(* IEC 61131-3 sources: brOscatLib/oscatBasic (part 2) *)

(* ---- DWORD_TO_STRB.st ---- *)
FUNCTION DWORD_TO_STRB
    (*http://www.oscat.de/images/OSCATBasic/oscat_basic333_en.pdf#page=153*)
    (* pointer für die ausgabe ermitteln *)
    pt ACCESS ADR(RETVAL);
    (* die 8 ausgabecharacter ermitteln und schreiben *)
    FOR i := 1 TO 32 DO
    	pt:= USINT_TO_BYTE(BOOL_TO_USINT(IN.31) + 48);
    	IN := SHL(IN,1);
    	pt ACCESS (ADR(pt) + 1);
    END_FOR

    (* der ausgabestring muss nochg mit 0 abgeschlossen werden *)
    pt := 0;
    DWORD_TO_STRB := TRUE;

    (* revision history
    hm		9.6.2007	rev 1.0
    	original version

    hm		15.dec 2007	rev 1.1
    	changed code for better performance

    hm	29. mar. 2008	rev 1.2
    	changed STRING to STRING(32)

    hm	20. jun. 2008	rev 1.3
    	performance improvement

    *)

END_FUNCTION

(* ---- DWORD_TO_STRF.st ---- *)
FUNCTION DWORD_TO_STRF
    (*http://www.oscat.de/images/OSCATBasic/oscat_basic333_en.pdf#page=154*)
    (* limit N to max 20 characters *)
    (* convert dword to string first and cut to length N *)
    temp := DWORD_TO_STRING(IN);
    FIX(temp,LIMIT(0,N,20),48,1, RETVAL);
    DWORD_TO_STRF := TRUE;

    (* revision history
    hm	26. jan.2007	rev 1.0
    	original version

    hm	29. mar. 2008	rev 1.1
    	changed STRING to STRING(20)
    	limit the output string to max 20 digits
    *)

END_FUNCTION

(* ---- DWORD_TO_STRH.st ---- *)
FUNCTION DWORD_TO_STRH
    (*http://www.oscat.de/images/OSCATBasic/oscat_basic333_en.pdf#page=154*)
    (* read output adress to pointer *)
    pt ACCESS (ADR(DWORD_TO_STRH) + 8);
    (* wirte the closing byte for the string *)
    pt:= 0;

    (* write the 8 hex characters backwards *)
    FOR i := 1 TO 8 DO;
    	(* decrement the pointer *)
    	pt ACCESS (ADR(pt) - 1);
    	(* read the lowest order hex value *)
    	temp := DWORD_TO_BYTE(IN AND 16#0000000F);
        intTemp := BYTE_TO_USINT(temp);
    	(* convert value to hex character *)
    	IF intTemp <= 9 THEN temp := USINT_TO_BYTE(intTemp + 48); ELSE temp := USINT_TO_BYTE(intTemp + 55); END_IF
    	(* write character to output string *)
    	pt := temp;
    	(* shift IN for nect hex character *)
    	IN := SHR(IN,4);
    END_FOR

    (* code beofre rev 1.2
    FOR i := 1 TO 8 DO
    	X := DWORD_TO_BYTE(IN AND 2#1111);
    	IF X <= 9 THEN X := X + 48; ELSE X := X + 55; END_IF
    	Cx := CHR(X);
    	temp := CONCAT(Cx, temp);
    	IN := SHR(IN,4);
    END_FOR
    DWORD_TO_STRH := temp;
    *)

    (* revision history
    hm	9. jun. 2007	rev 1.0
    	original version

    hm	11. sep. 2007	rev 1.1
    	changed coding for compatibility with twincat, concat cannot support a function as an argument.

    hm	15. dec. 2007	rev 1.2
    	changed code for better performance

    hm	29. mar. 2008	rev 1.3
    	changed STRING to STRING(8)

    *)

END_FUNCTION

(* ---- EASTER.st ---- *)
FUNCTION EASTER
    (*http://www.oscat.de/images/OSCATBasic/oscat_basic333_en.pdf#page=122*)
    b := (204 - 11 * (YEAR MOD 19)) MOD 30;
    IF b > 27 THEN b := b - 1; END_IF
    c := (YEAR + SHR(YEAR,2) + b - 13) MOD 7;
    oday := 28 + b - c;
    IF oday > 33 THEN
    	EASTER := SET_DATE(YEAR, 4, oday - 31);
    ELSE
    	EASTER := SET_DATE(YEAR, 3, oday);
    END_IF

    (* alternativer algorithmus ueber das pasah fest
    execution time roughly 200us
    Der sog. Passah-Vollmond wird berechnet, in dem das Jahr durch 19 ge-
    teilt wird und der Rest mit der folgenden Tabelle verglichen wird:

        0: Apr 14       5: Apr 18      10: Mrz 25      15: Mrz 30
        1: Apr 03       6: Apr 08      11: Apr 13      16: Apr 17
        2: Mrz 23       7: Mrz 28      12: Apr 02      17: Apr 07
        3: Apr 11       8: Apr 16      13: Mrz 22      18: Mrz 27
        4: Mrz 31       9: Apr 05      14: Apr 10

    Faellt dieses Datum auf einen Sonntag, ist Ostern der naechste Sonntag!

    Beispiel: 1992 MOD 19 = 16, daraus folgt 17.04., der naechste Sonntag
              ist dann der 19. April (Ostersonntag)
    *)

    (* this algorithm is 180 us
    a := YEAR MOD 19;
    b := YEAR / 100;
    c := YEAR MOD 100;
    d := b / 4;
    e := b MOD 4;
    f := (b + 8) / 25;
    g := (b - f + 1) / 3;
    h := (19 * a + b - d -g + 15) MOD 30;
    i := c / 4;
    k := c MOD 4;
    l := (32 + 2*e + 2*i - h - k) MOD 7;
    m := (a + 11 * h + 22 * l) / 451;
    x := h + l - 7 * m + 114;
    n := X / 31;
    o := x MOD 31 + 1;

    EASTER := set_Date(YEAR,n,o);
    *)
    (*
    Im Magazin "Nature" vom 20. April 1876 veröffentlichte ein anonymer Autor eine Tabelle mit Regeln zur Berechnung des (Gregorianischen) Ostersonntages des Jahres J. In Formeln ausgedrückt erhält man das Folgende:
    a	=	J mod 19
    b	=	int(J / 100)
    c	=	J mod 100
    d	=	int(b / 4)
    e	=	b mod 4
    f	=	int((b + 8) / 25)
    g	=	int((b - f + 1) / 3
    h	=	(19 · a + b - d - g + 15) mod 30
    i	=	int(c / 4)
    k	=	c mod 4
    l	=	(32 + 2 · e + 2 · i - h - k) mod 7
    m	=	int((a + 11 · h + 22 · l) / 451)
    n	=	int((h + l - 7 · m + 114) / 31)
    o	=	(h + l - 7 · m + 114) mod 31

    n ist hierbei die Nummer des Monats, o + 1 die Nummer des Tages auf welchen der Ostersonntag im Jahr J fällt. Dieser Algorithmus kommt ohne Hilfszahlen aus.

    *)

    (* revision history
    hm	27. dec 2006	rev 1.0
    	original version

    hm	15. dec 2007	rev 1.1
    	modified code for better performance

    hm	3. feb 2008		rev 1.2
    	modified code for better performance

    hm	7. apr. 2008	rev 1.3
    	improved performance
    *)
END_FUNCTION

(* ---- ELLIPSE_A.st ---- *)
FUNCTION ELLIPSE_A
    (*http://www.oscat.de/images/OSCATBasic/oscat_basic333_en.pdf#page=105*)
    ELLIPSE_A := cPI * R1 * R2;

    (* revision histroy
    hm	16. oct 2007	rev 1.0
    	original version

    hm	18. oct. 2008	rev 1.1
    	using math constants
    *)
END_FUNCTION

(* ---- ELLIPSE_C.st ---- *)
FUNCTION ELLIPSE_C
    (*http://www.oscat.de/images/OSCATBasic/oscat_basic333_en.pdf#page=106*)
    ELLIPSE_C := cPI * (3.0 * (R1+R2) - SQRT((3.0 * R1 + R2) * (3.0 * R2 + R1)));

    (* revision histroy
    hm	16. oct 2007	rev 1.0
    	original version

    hm	18. oct. 2008	rev 1.1
    	using math constants

    hm	10. mar. 2009	rev 1.2
    	changed syntax of real constants to 0.0

    *)
END_FUNCTION

(* ---- ERF.st ---- *)
FUNCTION ERF
    (*http://www.oscat.de/images/OSCATBasic/oscat_basic333_en.pdf#page=47*)
    x2 := X*X;
    ax2 := 0.147 * x2 + 1.0;
    ERF := SQRT(1.0 - EXP(-x2 * ((0.27323954473516 + ax2)/(ax2)))) * SGN(X);

    (* revision history
    hm	7. apr. 2008	rev 1.0
    	original version

    hm	30. jun. 2008	rev 1.1
    	added type conversions to avoid warnings under codesys 3.0

    hm	25. oct. 2008	rev 1.2
    	new code using new algorithm

    hm	10. mar. 2009	rev 1.3
    	real constants updated to new systax using dot
    *)
END_FUNCTION

(* ---- ERFC.st ---- *)
FUNCTION ERFC
    (*http://www.oscat.de/images/OSCATBasic/oscat_basic333_en.pdf#page=48*)
    ERFC := 1.0 - ERF(X);

    (* revision history
    hm	7. apr. 2008	rev 1.0
    	original version

    hm	10. mar. 2009	rev 1.1
    	real constants updated to new systax using dot

    *)
END_FUNCTION

(* ---- EVEN.st ---- *)
FUNCTION EVEN
    (*http://www.oscat.de/images/OSCATBasic/oscat_basic333_en.pdf#page=48*)
    EVEN := NOT IN.0;

    (* revision history
    hm	1. oct 2006	rev 1.0
    	ORIGINAL VERSION

    hm	01.12.2007	rev 1.1
    	changed code for improved performance

    hm	21. mar. 2008	rev 1.2
    	changed type of input IN from INT to DINT
    *)
END_FUNCTION

(* ---- EXEC.st ---- *)
FUNCTION EXEC
    (*http://www.oscat.de/images/OSCATBasic/oscat_basic333_en.pdf#page=155*)
    (* extract both numbers and operator *)
    TRIM(STR, temp);
    UPPERCASE(temp, RETVAL);

    pos := FINDB_NONUM(RETVAL);
    IF pos > 1 THEN R1 := STRING_TO_REAL(LEFT(RETVAL,pos-1)); END_IF
    R2 := STRING_TO_REAL(RIGHT(RETVAL,LEN(RETVAL)-pos));
    RETVAL := LEFT(RETVAL,pos);
    pos := FINDB_NUM(RETVAL);
    operator := RIGHT(RETVAL,LEN(RETVAL) - pos);
    IF operator = '' AND LEN(STR) = 0 THEN
    	RETVAL := '';
    	RETURN;
    ELSIF operator = '' THEN
    	RETVAL := STR;
    	RETURN;
    END_IF
    IF operator = '' THEN
    	RETVAL := REAL_TO_STRING(EXPT(R1, R2));
    ELSIF operator = 'SQRT' THEN
    	RETVAL := REAL_TO_STRING(SQRT(R2));
    ELSIF operator = 'SIN' THEN
    	RETVAL := REAL_TO_STRING(SIN(R2));
    ELSIF operator = 'COS' THEN
    	RETVAL := REAL_TO_STRING(COS(R2));
    ELSIF operator = 'TAN' THEN
    	RETVAL := REAL_TO_STRING(TAN(R2));
    ELSIF operator = '*' THEN
    	RETVAL := REAL_TO_STRING(R1 * R2);
    ELSIF operator = '/' THEN
    	IF R2 <> 0 THEN RETVAL := REAL_TO_STRING(R1 / R2); ELSE RETVAL := 'ERROR'; END_IF
    ELSIF operator = '+' THEN
    	RETVAL := REAL_TO_STRING(R1 + R2);
    ELSIF operator = '-' THEN
    	RETVAL := REAL_TO_STRING(R1 - R2);
    ELSE
    	RETVAL := 'ERROR';
    END_IF

    IF RETVAL = 'ERROR' THEN
        EXEC := FALSE;
    	RETURN;
    (* some systems deliver integer instead of real *)
    ELSIF FIND(RETVAL,'.') = 0 THEN
    	RETVAL := CONCAT(RETVAL, '.0');
    (* some systems deliver n. instead of n.0 ! *)
    ELSIF RIGHT(RETVAL,1) = '.' THEN
    	RETVAL := CONCAT(RETVAL,'0');
    END_IF
    EXEC := TRUE;

    (* revision history

    hm 	6.feb 2007		rev 1.1
    	cos has to be written in uppercase
    	divide by 0 will return an error

    hm	5. mar. 2008	rev 1.2
    	add a 0 to the string if a '.' is at the end of the string

    hm	20. mar. 2008	rev 1.3
    	make sure the function always returns a real value in the form of x.y

    hm	29. mar. 2008	rev 1.4
    	changed STRING to STRING(STRING_LENGTH)
    *)
END_FUNCTION

(* ---- EXP10.st ---- *)
FUNCTION EXP10
    (*http://www.oscat.de/images/OSCATBasic/oscat_basic333_en.pdf#page=49*)
    EXP10 := EXP(X * 2.30258509299405);

    (* revision history
    hm	2. dec 2007		rev 1.0
    	original version

    *)
END_FUNCTION

(* ---- EXPN.st ---- *)
FUNCTION EXPN
    (*http://www.oscat.de/images/OSCATBasic/oscat_basic333_en.pdf#page=49*)
    sign := N.15;
    N := ABS(N);
    IF N.0 THEN EXPN := X; ELSE EXPN := 1.0; END_IF
    N := SHR(N,1);
    WHILE N > 0 DO
       X := X * X;
       IF N.0 THEN EXPN := EXPN * X; END_IF
       N := SHR(N,1);
    END_WHILE
    IF sign THEN EXPN := 1.0 / EXPN; END_IF

    (* revision history
    hm	4. dec 2007	rev 1.0
    	original version

    hm	22. oct. 2008	rev 1.1
    	optimized code

    hm	10. mar. 2009	rev 1.2
    	removed nested comments
    	real constants updated to new systax using dot

    *)
END_FUNCTION

(* ---- F_LIN.st ---- *)
FUNCTION F_LIN
    (*http://www.oscat.de/images/OSCATBasic/oscat_basic333_en.pdf#page=96*)
    F_LIN := A * X + B;

END_FUNCTION

(* ---- F_LIN2.st ---- *)
FUNCTION F_LIN2
    (*http://www.oscat.de/images/OSCATBasic/oscat_basic333_en.pdf#page=96*)
    F_LIN2 := (Y2 - Y1) / (X2 - X1) * (X - X1) + Y1;

    (* revision history
    hm	1. jan. 2007	rev 1.0
    	original release

    hm	17. dec. 2008	rev 1.1
    	optimized formula

    *)
END_FUNCTION

(* ---- F_POLY.st ---- *)
FUNCTION F_POLY
    (*http://www.oscat.de/images/OSCATBasic/oscat_basic333_en.pdf#page=97*)
    F_POLY := ((((((( C[7] * X + C[6] ) * X + C[5] ) * X + C[4] ) * X + C[3] ) * X + C[2] ) * X + C[1] ) * X + C[0] ) ;

    (* revision history
    hm		20. may. 2008		rev 1.0
    	original version

    hm	18. mar. 2011	rev 1.1
    	improved performance
    *)

END_FUNCTION

(* ---- F_POWER.st ---- *)
FUNCTION F_POWER
    (*http://www.oscat.de/images/OSCATBasic/oscat_basic333_en.pdf#page=97*)
    F_POWER := A * EXPT(X, N);

END_FUNCTION

(* ---- F_QUAD.st ---- *)
FUNCTION F_QUAD
    (*http://www.oscat.de/images/OSCATBasic/oscat_basic333_en.pdf#page=97*)
    F_QUAD :=  (A * X + B) * X + C;

    (* revision history

    hm	1. sep. 2006	rev 1.0
    	original version

    hm	18. mar. 2001	rev 1.1
    	improved performance
    *)
END_FUNCTION

(* ---- F_TO_C.st ---- *)
FUNCTION F_TO_C
    (*http://www.oscat.de/images/OSCATBasic/oscat_basic333_en.pdf#page=361*)
    F_TO_C := (FAHRENHEIT - 32.0) * 0.5555555555555;

    (* revision history
    hm	4. aug 2006	rev 1.0
    	original version

    hm	11. mar. 2009	rev 1.1
    	real constants updated to new systax using dot

    *)
END_FUNCTION

(* ---- F_TO_OM.st ---- *)
FUNCTION F_TO_OM
    (*http://www.oscat.de/images/OSCATBasic/oscat_basic333_en.pdf#page=362*)
    F_TO_OM := cPI2 * F;

    (* revision history
    hm	22. jan. 2007	rev 1.0
    	original version

    hm	18. oct. 2008	rev 1.1
    	unsing math constants

    *)
END_FUNCTION

(* ---- F_TO_PT.st ---- *)
FUNCTION F_TO_PT
    (*http://www.oscat.de/images/OSCATBasic/oscat_basic333_en.pdf#page=362*)
    F_TO_PT := DWORD_TO_TIME(REAL_TO_DWORD(1.0 / F * 1000.0));

    (* revision history

    hm	4. aug. 2006	rev 1.0
    	original version

    hm	11. mar. 2009	rev 1.1
    	real constants updated to new systax using dot

    *)

END_FUNCTION

(* ---- FACT.st ---- *)
FUNCTION FACT
    (*http://www.oscat.de/images/OSCATBasic/oscat_basic333_en.pdf#page=49*)
    IF X >= 0 AND X <= 12 THEN
    	FACT := cFACTS[X];
    ELSE
    	FACT := -1;
    END_IF

    (* working code without array
    IF X > 12 OR X < 0 THEN
    	FACT := -1;
    ELSIF X < 7 THEN
    	FACT := 1;
    	FOR i := 2 TO X DO
    		FACT := FACT * i;
    	END_FOR
    ELSE
    	FACT := 5040;
    	FOR i := 8 TO X DO
    		FACT := FACT * i;
    	END_FOR
    END_IF
    *)

    (* revision history
    hm 4.3.2007		rev 1.1
    	changed a critical error where while loop was indefinite.

    hm	10.12.2007	rev 1.2
    	start value for i has changed to 2 for better performance

    hm	10. mar 2008	rev 1.3
    	changed output of FACT to dint to allow bigger values

    hm	27. oct. 2008	rev 1.4
    	optimized code

    hm	26. mar. 2011	rev 1.5
    	using array cfacts
    *)
END_FUNCTION

(* ---- FIB.st ---- *)
FUNCTION FIB
    (*http://www.oscat.de/images/OSCATBasic/oscat_basic333_en.pdf#page=50*)
    IF X < 0 OR X > 46 THEN
    	FIB := -1;
    ELSIF X < 2 THEN
    	FIB := X;
    	RETURN;
    ELSE
    	(* the fibonacci number is the sum of the two suceeding fibonaci numbers *)
    	(* we store the numbers alternatively in t1 and t2 depending on pt *)
    	t2 := 1;
    	WHILE X > 3 DO
    		X := X-2;
    		t1 := t1 + t2;
    		t2 := t1 + t2;
    	END_WHILE
    	IF X > 2 THEN t1 := t1 + t2; END_IF
    	FIB := t1 + t2;
    END_IF

    (* alternative code for very big numbers

    IF X < 31 THEN
    	FIB := 0.4472136 * (expn(1.618034,X) - expn(-0.618034,X));
    ELSE
    	FIB := 0.4472133 * expn(1.618034,X);
    END_IF

    *)

    (* revision history
    hm		27. dec 2007	rev 1.0
    	original version

    hm		2. jan 2008	rev 1.1
    	deleted unused variable pt

    hm		10. mar 2008	rev 1.2
    	changed output to dint instead of real

    hm		26. mar. 2008	rev 1.3
    	function now returns -1 for input < 0 or > 46

    *)
END_FUNCTION

(* ---- FILL.st ---- *)
FUNCTION FILL
    (*http://www.oscat.de/images/OSCATBasic/oscat_basic333_en.pdf#page=155*)
    CHR_TO_STRING(C, sx);
    (* limit L to maximum 80 characters the length of a standard string *)
    L := LIMIT(0,L,STRING_LENGTH);
    (* create a string of characters to be connected to str *)
    FOR i := 1 TO 8 DO
    	RETVAL := CONCAT(RETVAL,RETVAL);
    	IF L.7 THEN RETVAL := CONCAT(RETVAL,sx); END_IF
    	L := SHL(L,1);
    END_FOR
    FILL:=TRUE;

    (* revision histroy
    hm	29. mar. 2008	rev 1.0
    	original release

    hm	17. dec. 2008	rev 1.1
    	changed function chr to chr_to_string

    *)
END_FUNCTION

(* ---- FIND_CHAR.st ---- *)
FUNCTION FIND_CHAR
    (*http://www.oscat.de/images/OSCATBasic/oscat_basic333_en.pdf#page=156*)
    pt ACCESS ADR(STR);
    stop := LEN(STR);
    FOR i := MAX(POS,1) TO stop DO;
    	X := pt[i];
    	IF X > 31 AND ((cEXTENDED_ASCII AND X <> 127) OR (NOT cEXTENDED_ASCII AND X < 127)) THEN
    		FIND_CHAR := i;
    		RETURN;
    	END_IF
    END_FOR
    FIND_CHAR := 0;

    (* revision history
    hm	29. feb 2008	rev 1.0
    	original version

    hm	26. mar. 2008	rev 1.1
    	char will now accept extended ascii

    hm	29. mar. 2008	rev 1.2
    	changed STRING to STRING(STRING_LENGTH)

    hm	21. oct. 2008	rev 1.3
    	changes setup constants
    	optimized code
    *)

END_FUNCTION

(* ---- FIND_CTRL.st ---- *)
FUNCTION FIND_CTRL
    (*http://www.oscat.de/images/OSCATBasic/oscat_basic333_en.pdf#page=157*)
    pt ACCESS ADR(STR);
    stop := LEN(STR);
    FOR i := MAX(POS,1) TO stop DO;
    	x := pt[i];
    	IF x < 32 OR x = 127 THEN
    		FIND_CTRL := i;
    		RETURN;
    	END_IF
    END_FOR
    FIND_CTRL := 0;

    (* revision history
    hm	29. feb 2008	rev 1.0
    	original version

    hm	26. mar. 2008	rev 1.1
    	character 127 is now recognized as control

    hm	29. mar. 2008	rev 1.2
    	changed STRING to STRING(STRING_LENGTH)
    *)
END_FUNCTION

(* ---- FIND_NONUM.st ---- *)
FUNCTION FIND_NONUM
    (*http://www.oscat.de/images/OSCATBasic/oscat_basic333_en.pdf#page=157*)
    pt ACCESS ADR(STR);
    end := LEN(STR);
    FOR i := MAX(POS,1) TO end DO;
    	X := pt[i];
    	IF (X < 48 AND X <> 46) OR X > 57 THEN
    		FIND_NONUM := i;
    		RETURN;
    	END_IF
    END_FOR
    FIND_NONUM := 0;

    (* revision history
    hm	6. oct. 2006	rev 1.0
    	original version

    hm	29. feb 2008	rev 1.1
    	added input POS to start search at position

    hm	29. mar. 2008	rev 1.2
    	changed STRING to STRING(STRING_LENGTH)

    hm	21. oct. 2008	rev 1.3
    	optimized code

    *)
END_FUNCTION

(* ---- FIND_NUM.st ---- *)
FUNCTION FIND_NUM
    (*http://www.oscat.de/images/OSCATBasic/oscat_basic333_en.pdf#page=157*)
    pt ACCESS ADR(STR);
    stop := LEN(STR);
    FOR i := MAX(POS,1) TO stop DO;
    	X := pt[i];
    	IF (X > 47 AND X < 58) OR X = 46 THEN
    		FIND_NUM := i;
    		RETURN;
    	END_IF
    END_FOR
    FIND_NUM := 0;

    (* revision history
    hm	6. oct. 2006	rev 1.0
    	original version

    hm	29. feb 2008	rev 1.1
    	added input POS to start search at position

    hm	29. mar. 2008	rev 1.2
    	changed STRING to STRING(STRING_LENGTH)

    *)
END_FUNCTION

(* ---- FINDB.st ---- *)
FUNCTION FINDB
    (*http://www.oscat.de/images/OSCATBasic/oscat_basic333_en.pdf#page=158*)
    length := LEN(STR2);
    FOR pos := LEN(STR1) - length + 1 TO 1 BY -1 DO
    	IF MID(STR1,length,pos) = STR2 THEN
    		FINDB := pos;
    		RETURN;
    	END_IF
    END_FOR
    FINDB := 0;

    (* revision history
    hm	6. oct 2006		rev 1.0
    	original version

    hm	15 dec 2007		rev 1.1
    	changed code for better performance

    hm	29. feb 2008	rev 1.2
    	added FINDB := 0 for compatibility reasons

    hm	29. mar. 2008	rev 1.3
    	changed STRING to STRING(STRING_LENGTH)
    *)
END_FUNCTION

(* ---- FINDB_NONUM.st ---- *)
FUNCTION FINDB_NONUM
    (*http://www.oscat.de/images/OSCATBasic/oscat_basic333_en.pdf#page=158*)
    pt ACCESS (ADR(STR) + LEN(STR) - 1);
    FOR pos := LEN(STR) TO 1 BY -1 DO;
    	IF (pt < 48 AND pt <> 46) OR pt > 57 THEN
    		FINDB_NONUM := pos;
    		RETURN;
    	END_IF
    	pt ACCESS (ADR(pt) - 1);
    END_FOR
    FINDB_NONUM := 0;

    (* revision history
    hm	6. oct 2006		rev 1.0
    	original version

    hm	29. feb 2008	rev 1.1
    	improved performance

    hm	29. mar. 2008	rev 1.2
    	changed STRING to STRING(STRING_LENGTH)

    hm	21. oct. 2008	rev 1.3
    	optimized code
    *)
END_FUNCTION

(* ---- FINDB_NUM.st ---- *)
FUNCTION FINDB_NUM
    (*http://www.oscat.de/images/OSCATBasic/oscat_basic333_en.pdf#page=159*)
    pt ACCESS (ADR(STR) + LEN(STR) - 1);
    FOR pos := LEN(STR) TO 1 BY -1 DO;
    	IF (pt > 47 AND pt < 58) OR pt = 46 THEN
    		FINDB_NUM := pos;
    		RETURN;
    	END_IF
    	pt ACCESS (ADR(pt) - 1);
    END_FOR
    FINDB_NUM := 0;

    (* revision history
    hm	6. oct 2006		rev 1.0
    	original version

    hm	29. feb 2008	rev 1.1
    	improved performance

    hm	29. mar. 2008	rev 1.2
    	changed STRING to STRING(STRING_LENGTH)
    *)
END_FUNCTION

(* ---- FINDP.st ---- *)
FUNCTION FINDP
    (*http://www.oscat.de/images/OSCATBasic/oscat_basic333_en.pdf#page=159*)
    ls := LEN(STR);
    lx := LEN(SRC);
    IF ls < lx OR lx = 0 THEN RETURN; END_IF
    stp := ls - lx + 1;
    FOR i := MAX(POS,1) TO stp DO
    	IF MID(STR,lx,i) = SRC THEN
    		FINDP := i;
    		RETURN;
    	END_IF
    END_FOR
    FINDP := 0;

    (* revision histroy
    hm	4. feb. 2008	rev 1.0
    	original release

    hm	29. feb 2008	rev 1.1
    	ADDED MAX(POS,1) in loop initialization

    hm	29. mar. 2008	rev 1.2
    	changed STRING to STRING(STRING_LENGTH)
    *)

END_FUNCTION

(* ---- FIX.st ---- *)
FUNCTION FIX
    (*http://www.oscat.de/images/OSCATBasic/oscat_basic333_en.pdf#page=160*)
    (* make sure L does not exceed the limits of a string *)
    N := LIMIT(0,L,STRING_LENGTH) - LEN(STR);
    IF N <= 0 THEN
    	(* truncate the string at length N *)
    	IF M = 1 THEN
    		RETVAL := RIGHT(STR,L);
    	ELSE
    		RETVAL := LEFT(STR,L);
    	END_IF
    ELSIF M = 1 THEN
    	(* connect fill characters at the beginning *)
    	FILL(C,N, SX);
    	RETVAL := CONCAT(SX,STR);
    ELSIF M = 2 THEN
    	(* center STR beween fill characters *)
    	(* for an uneven number of fill characters, there is one more at the end *)
    	FILL(C,SHR(N+1,1), SX);
    	RETVAL := CONCAT(STR,SX);
    	SX := LEFT(SX,SHR(N,1));
    	RETVAL := CONCAT(SX,RETVAL);
    ELSE
    	(* connect fill characters at the end *)
    	FILL(C,N, SX);
    	RETVAL := CONCAT(STR,SX);
    END_IF
    FIX := TRUE;

    (* revision histroy
    hm	29. mar. 2008	rev 1.0
    	original release

    *)
END_FUNCTION

(* ---- FLOAT_TO_REAL.st ---- *)
FUNCTION FLOAT_TO_REAL
    (*http://www.oscat.de/images/OSCATBasic/oscat_basic333_en.pdf#page=160*)
    pt ACCESS ADR(FLT);
    stop := LEN(FLT);

    (* we first check for sign and exit if first number or dot is reached *)
    FOR i := 1 TO stop DO
    	X := pt[i];
        intX := BYTE_TO_USINT(X);
    	IF intX > 47 AND intX < 58 OR intX = 46 THEN
    		EXIT;
    	ELSIF intX = 45 THEN
    		(* code 45 is sign *)
    		sign := -1;
    	END_IF
    END_FOR

    (* now we scan numbers till end or dot or E is reached *)
    FOR i := i TO stop DO
    	X := pt[i];
        intX := BYTE_TO_USINT(X);
    	IF intX = 44 OR intX = 46 OR intX = 69 OR intX = 101 THEN
    		EXIT;
    	(* calculate the value of the digit *)
    	ELSIF intX > 47 AND intX < 58 THEN
    		tmp := tmp * 10 + intX - 48;
    	END_IF
    END_FOR

    (* process the portion after the comma if comma or dot is reached exit if exponent starts *)
    IF X = 44 OR X = 46 THEN
    	FOR i := i + 1 TO stop DO
    		X := pt[i];
            intX := BYTE_TO_USINT(X);
    		IF intX = 69 OR intX = 101 THEN
    			EXIT;
    		ELSIF intX > 47 AND intX < 58 THEN
    			tmp := tmp * 10 + intX - 48;
    			d := d - 1;
    		END_IF
    	END_FOR
    END_IF

    (* process exponent if present *)
    IF intX = 69 OR intX = 101 THEN
    	d := d + DEC_TO_INT(RIGHT(FLT, stop - i));
    END_IF

    FLOAT_TO_REAL :=  EXPN(10, d) * DINT_TO_REAL(tmp * sign);

    (* revision histroy
    hm	22. jun. 2008	rev 1.0
    	original release

    hm	2. oct. 2008	rev 1.1
    	fixed an error, characters 8 and 9 would not be converted

    hm	22. oct. 2008	rev 1.2
    	last fix was not done correctly

    hm	23. oct. 2008	rev 1.3
    	optimzed code
    *)

END_FUNCTION

(* ---- FLOOR.st ---- *)
FUNCTION FLOOR
    (*http://www.oscat.de/images/OSCATBasic/oscat_basic333_en.pdf#page=50*)
    FLOOR := REAL_TO_INT(X);
    IF FLOOR > X THEN
    	FLOOR := FLOOR - 1;
    END_IF

    (* revision history
    hm		7. feb 2007		rev 1.0
    	originlal version

    hm		21. mar. 2008	rev 1.1
    	replaced trunc with real_to_int for compatibility reasons

    *)
END_FUNCTION

(* ---- FLOOR2.st ---- *)
FUNCTION FLOOR2
    (*http://www.oscat.de/images/OSCATBasic/oscat_basic333_en.pdf#page=51*)
    FLOOR2 := REAL_TO_DINT(X);
    IF DINT_TO_REAL(FLOOR2) > X THEN
    	FLOOR2 := FLOOR2 - 1;
    END_IF

    (* revision history
    hm	21. mar. 2008	rev 1.0
    	originlal version

    hm	4. apr. 2008	rev 1.1
    	added type conversion to avoid warnings under codesys 3.0
    *)
END_FUNCTION

(* ---- FRACT.st ---- *)
FUNCTION FRACT
    (*http://www.oscat.de/images/OSCATBasic/oscat_basic333_en.pdf#page=51*)
    IF ABS(X) < 2.0E9 THEN
    	FRACT := X - DINT_TO_REAL(D_TRUNC(X));
    ELSE
    	FRACT := 0.0;
    END_IF

    (* revision history
    hm	4. aug 2006	rev 1.0
    	original version

    hm	11. mar 2008	rev 1.1
    	added dint_to_real for compatibility reasons
    	now returns 0 for number > 2e9
    	changed input to X

    hm	21. mar. 2008	rev 1.2
    	use D_trunc instead of TRUNC for compatibility reasons

    hm	10. mar. 2009	rev 1.3
    	real constants updated to new systax using dot

    *)
END_FUNCTION

(* ---- FRMP_B.st ---- *)
FUNCTION FRMP_B
    (*http://www.oscat.de/images/OSCATBasic/oscat_basic333_en.pdf#page=98*)
    IF TD < TR THEN
    	FRMP_B := USINT_TO_BYTE(MIN(UDINT_TO_USINT(SHL(TIME_TO_UDINT(TD), 8) / TIME_TO_UDINT(TR)), SEL(DIR, BYTE_TO_USINT(START), 255 - BYTE_TO_USINT(START))));
    	IF DIR THEN
    		FRMP_B := USINT_TO_BYTE(BYTE_TO_USINT(START) + BYTE_TO_USINT(FRMP_B));
    	ELSE
    		FRMP_B := USINT_TO_BYTE(BYTE_TO_USINT(START) - BYTE_TO_USINT(FRMP_B));
    	END_IF
    ELSE
    	FRMP_B := SEL(DIR, BYTE#0, BYTE#255);
    END_IF

    (* revision history

    17. feb. 2011	rev 1.0
    	new module

    *)
END_FUNCTION

(* ---- FSTRING_TO_BYTE.st ---- *)
FUNCTION FSTRING_TO_BYTE
    (*http://www.oscat.de/images/OSCATBasic/oscat_basic333_en.pdf#page=161*)
    IF LEFT(IN, 2) = '2#' THEN
    	(* we need to convert binary *)
    	FSTRING_TO_BYTE := BIN_TO_BYTE(RIGHT(IN, LEN(IN) - 2));
    ELSIF LEFT(IN, 2) = '8#' THEN
    	(* weneed to convert octals *)
    	FSTRING_TO_BYTE := OCT_TO_BYTE(RIGHT(IN, LEN(IN) - 2));
    ELSIF LEFT(IN, 3) = '16#' THEN
    	(* we need to convert hexadecimal *)
    	FSTRING_TO_BYTE := HEX_TO_BYTE(RIGHT(IN, LEN(IN) - 3));
    ELSE
    	(* we assume decimal representation *)
        CLEAN(IN,'0123456789', temp);
    	FSTRING_TO_BYTE := DEC_TO_BYTE(temp);
    END_IF

    (* revision histroy
    hm	18. jun. 2008	rev 1.0
    	original release

    hm	20. sep. 2008	rev 1.1
    	changed length of input string from 20 to 12
    *)

END_FUNCTION

(* ---- FSTRING_TO_DT.st ---- *)
FUNCTION FSTRING_TO_DT
    (*http://www.oscat.de/images/OSCATBasic/oscat_basic333_en.pdf#page=161*)
    (* scan input string *)
    WHILE FMT <> '' DO
    	c := LEFT(FMT,1);
    	IF c = ignore THEN
    		(* skip ignore characters *)
    		FMT := DELETE(FMT,1,1);
    		SDT := DELETE(SDT,1,1);
    	ELSIF c = fchar THEN
    		(* format chracter found skip format char and read identifier *)
    		(* store format identifier in c and skip to next char in FMT *)
    		c := MID(FMT,1,2);
    		FMT := DELETE(FMT,2,1);
    		(* extract the substring until the end of SDT or to next char of FMT *)
    		IF FMT = '' THEN
    			tmp := SDT;
    		ELSE
    			(* serach for end of substring *)
    			end := FIND(SDT, LEFT(FMT,1))-1;
    			tmp := LEFT(SDT, end);
    			SDT := DELETE(SDT, end,1);
    		END_IF
    		(* extract information from substring *)
    		IF c = 'Y' THEN
    			dy := STRING_TO_INT(tmp);
    			IF dy < 100 THEN dy := dy + 2000; END_IF
    		ELSIF c = 'M' THEN
    			dm := STRING_TO_INT(tmp);
    		ELSIF c = 'N' THEN
    			dm := FSTRING_TO_MONTH(tmp,0);
    		ELSIF c = 'D' THEN
    			dd := STRING_TO_INT(tmp);
    		ELSIF c = 'h' THEN
    			th := STRING_TO_INT(tmp);
    		ELSIF c = 'm' THEN
    			tm := STRING_TO_INT(tmp);
    		ELSIF c = 's' THEN
    			ts := STRING_TO_INT(tmp);
    		END_IF
    	ELSIF c = LEFT(SDT,1) THEN
    		(* skip matching characters *)
    		FMT := DELETE(FMT,1,1);
    		SDT := DELETE(SDT,1,1);
    	ELSE
    		RETURN;
    	END_IF
    END_WHILE

    FSTRING_TO_DT := SET_DT(dy,dm,dd,th,tm,ts);

    (* revision histroy
    hm	24. sep. 2008	rev 1.0
    	original release

    *)

END_FUNCTION

(* ---- FSTRING_TO_DWORD.st ---- *)
FUNCTION FSTRING_TO_DWORD
    (*http://www.oscat.de/images/OSCATBasic/oscat_basic333_en.pdf#page=162*)
    IF LEFT(IN, 2) = '2#' THEN
    	(* we need to convert binary *)
    	FSTRING_TO_DWORD := BIN_TO_DWORD(RIGHT(IN, LEN(IN) - 2));
    ELSIF LEFT(IN, 2) = '8#' THEN
    	(* weneed to convert octals *)
    	FSTRING_TO_DWORD := OCT_TO_DWORD(RIGHT(IN, LEN(IN) - 2));
    ELSIF LEFT(IN, 3) = '16#' THEN
    	(* we need to convert hexadecimal *)
    	FSTRING_TO_DWORD := HEX_TO_DWORD(RIGHT(IN, LEN(IN) - 3));
    ELSE
    	(* we assume decimal representation *)
        CLEAN(IN,'0123456789', temp);
    	FSTRING_TO_DWORD := DEC_TO_DWORD(temp);
    END_IF

    (* revision histroy
    hm	18. jun. 2008	rev 1.0
    	original release

    hm	20. sep. 2008	rev 1.1
    	changed length of input dtring from 20 to 40

    *)

END_FUNCTION

(* ---- FSTRING_TO_MONTH.st ---- *)
FUNCTION FSTRING_TO_MONTH
    (*http://www.oscat.de/images/OSCATBasic/oscat_basic333_en.pdf#page=162*)
    IF LANG = 0 THEN lx := cLANGUAGE_DEFAULT; ELSE lx := MIN(LANG, cLANGUAGE_LMAX); END_IF
    TRIM(MTH, MTH);
    LOWERCASE(MTH, MTH);
    CAPITALIZE(MTH, MTH);

    FOR FSTRING_TO_MONTH := 1 TO 12 DO
    	IF MTH = cMONTHS[lx, FSTRING_TO_MONTH] THEN RETURN; END_IF
    	IF MTH = cMONTHS3[lx, FSTRING_TO_MONTH] THEN RETURN; END_IF
    END_FOR

    (* since no name matched try to decode as integer *)
    FSTRING_TO_MONTH := STRING_TO_INT(MTH);

    (* revision histroy
    hm	25. sep. 2008	rev 1.0
    	original release

    hm	19. oct. 2008	rev 1.1
    	changed language setup constants

    hm	25. oct. 2008	rev 1.2
    	optimized code
    *)

END_FUNCTION

(* ---- FSTRING_TO_WEEK.st ---- *)
FUNCTION FSTRING_TO_WEEK
    (*http://www.oscat.de/images/OSCATBasic/oscat_basic333_en.pdf#page=163*)
    pos := FIND(WEEK, ',');
    WHILE pos > 0 DO
    	FSTRING_TO_WEEK := FSTRING_TO_WEEK OR SHR(BYTE#128, FSTRING_TO_WEEKDAY(MID(WEEK, pos - 1, 1), LANG));
    	WEEK := RIGHT(WEEK, LEN(WEEK) - pos);
    	pos := FIND(WEEK, ',');
    END_WHILE
    FSTRING_TO_WEEK := (FSTRING_TO_WEEK OR SHR(BYTE#128, FSTRING_TO_WEEKDAY(WEEK, LANG))) AND BYTE#127;

    (* revision histroy
    hm	18. jun. 2008	rev 1.0
    	original release

    hm	25. oct. 2008	rev 1.1
    	using language defauls and input LANG
    *)

END_FUNCTION

(* ---- FSTRING_TO_WEEKDAY.st ---- *)
FUNCTION FSTRING_TO_WEEKDAY
    (*http://www.oscat.de/images/OSCATBasic/oscat_basic333_en.pdf#page=164*)
    IF LANG = 0 THEN ly := cLANGUAGE_DEFAULT; ELSE ly := MIN(LANG, cLANGUAGE_LMAX); END_IF
    (* tmp needs to be calculated first otherwise find can return wrong values *)
    TRIM(WDAY, tmp);
    LOWERCASE(tmp, tmp);
    CAPITALIZE(tmp, tmp);
    FOR i := 1 TO 7 DO
    	IF cWEEKDAYS2[ly, i] = tmp THEN
    		FSTRING_TO_WEEKDAY := i;
    		RETURN;
    	END_IF
    END_FOR
    FSTRING_TO_WEEKDAY := STRING_TO_INT(WDAY);

    (* revision histroy
    hm	18. jun. 2008	rev 1.0
    	original release

    hm	18. jul. 2008	rev 1.1
    	changed nested call of left(trim()) for compatibility reasons

    hm	25. oct. 2008	rev 1.2
    	using language constants
    *)

END_FUNCTION

(* ---- GAMMA.st ---- *)
FUNCTION GAMMA
    (*http://www.oscat.de/images/OSCATBasic/oscat_basic333_en.pdf#page=52*)
    IF X > 0.0 THEN
    	GAMMA := SQRT(cPI2 / X) * EXPT(ce_INV * (X + 1.0 / (12.0 * X - 0.1 / X)), X);
    END_IF

    (* the stirling formula is not very accurate for small values of X
    IF X >=0 THEN GAMMA := SQRT(cPI2 * X) * EXPT(X / ce, X); END_IF
    *)

    (* revision history
    hm	10.12.2007	rev 1.0
    	original version

    hm	18. oct. 2008	rev 1.1
    	using math constants

    hm	26. oct. 2008	rev 1.2
    	using new formula with better accuracy

    hm	10. mar. 2009	rev 1.3
    	real constants updated to new systax using dot

    *)
END_FUNCTION

(* ---- GAUSS.st ---- *)
FUNCTION GAUSS
    (*http://www.oscat.de/images/OSCATBasic/oscat_basic333_en.pdf#page=52*)
    temp := X - U;
    si_inv := 1.0  / SI;
    GAUSS := EXP(temp * temp * si_inv * si_inv * - 0.5) * 0.39894228 * si_inv;

    (* revision hisdtory
    hm	6. apr. 2008	rev 1.0
    	original version

    hm	27. oct. 2008	rev 1.1
    	optimized performance

    hm	10. mar. 2009	rev 1.2
    	real constants updated to new systax using dot

    *)
END_FUNCTION

(* ---- GAUSSCD.st ---- *)
FUNCTION GAUSSCD
    (*http://www.oscat.de/images/OSCATBasic/oscat_basic333_en.pdf#page=53*)
    GAUSSCD := (ERF((X - U) / (SI * 1.414213562)) + 1.0) * 0.5;

    (* revision hisdtory
    hm	6. apr. 2008	rev 1.0
    	original version

    hm	10. mar. 2009	rev 1.1
    	real constants updated to new systax using dot

    *)
END_FUNCTION

(* ---- GCD.st ---- *)
FUNCTION GCD
    (*http://www.oscat.de/images/OSCATBasic/oscat_basic333_en.pdf#page=53*)
    IF A = 0 THEN
    	GCD := DINT_TO_INT(ABS(B));
    ELSIF B = 0 THEN
    	GCD := DINT_TO_INT(ABS(A));
    ELSE
    	A := ABS(A);
    	B := ABS(B);
    	GCD := 1;
    	WHILE NOT(A.0 OR B.0) DO
    		A := SHR(A,1);
    		B := SHR(B,1);
    		GCD := SHL(GCD,1);
    	END_WHILE
    	WHILE A > 0 DO
    		IF NOT(A.0) THEN A := SHR(A,1);
    		ELSIF NOT(B.0) THEN B := SHR(B,1);
    		ELSE
    			t:= SHR(ABS(A-B),1);
    			IF A < B THEN B := t; ELSE A := t; END_IF
    		END_IF
    	END_WHILE
    	GCD := GCD * DINT_TO_INT(B);
    END_IF

    (* revision history
    hm	19. jan. 2011	rev 1.0
    	original version

    *)
END_FUNCTION

(* ---- GDF.st ---- *)
FUNCTION GDF
    (*http://www.oscat.de/images/OSCATBasic/oscat_basic333_en.pdf#page=54*)
    IF X = 0.0 THEN
    	GDF := 0.0;
    ELSIF X > 15.0 THEN
    	GDF := cPI05;
    ELSIF X < -15.0 THEN
    	GDF := -cPI05;
    ELSE
    	GDF := ATAN(EXP(X)) * 2.0 - cPI05;
    END_IF

    (* revision history
    hm	27. apr. 2008	rev 1.0
    	original version

    hm	18. oct. 2008	rev 1.1
    	using math constants

    hm	10. mar. 2009	rev 1.2
    	real constants updated to new systax using dot

    *)

END_FUNCTION

(* ---- GEO_TO_DEG.st ---- *)
FUNCTION GEO_TO_DEG
    (*http://www.oscat.de/images/OSCATBasic/oscat_basic333_en.pdf#page=362*)
    GEO_TO_DEG := INT_TO_REAL(D) + INT_TO_REAL(M) * 0.016666666666667 + SEC * 0.00027777777777778;

    (* revision histroy
    hm	22. jan. 2009	rev 1.0
    	original release

    *)
END_FUNCTION

(* ---- GOLD.st ---- *)
FUNCTION GOLD
    (*http://www.oscat.de/images/OSCATBasic/oscat_basic333_en.pdf#page=54*)
    GOLD := (X + SQRT(X*X + 4.0)) * 0.5;

    (* revision history
    hm	27. apr. 2008	rev 1.0
    	original version

    hm	10. mar. 2009	rev 1.1
    	real constants updated to new systax using dot

    *)

END_FUNCTION

(* ---- GRAY_TO_BYTE.st ---- *)
FUNCTION GRAY_TO_BYTE
    (*http://www.oscat.de/images/OSCATBasic/oscat_basic333_en.pdf#page=226*)
    GRAY_TO_BYTE := SHR(IN,4) XOR IN;
    GRAY_TO_BYTE := SHR(GRAY_TO_BYTE,2) XOR GRAY_TO_BYTE;
    GRAY_TO_BYTE := SHR(GRAY_TO_BYTE,1) XOR GRAY_TO_BYTE;

    (* revision history
    hm	9. nov. 2009	rev 1.0
    	original version

    *)
END_FUNCTION

(* ---- HEX_TO_BYTE.st ---- *)
FUNCTION HEX_TO_BYTE
    (*http://www.oscat.de/images/OSCATBasic/oscat_basic333_en.pdf#page=164*)
    pt ACCESS ADR(HEX);
    stop := LEN(HEX);
    FOR i := 1 TO stop DO
    	(* read the first character and subtract 48 to get value in decimal 0 = 48 *)
    	X := pt;
        intX := BYTE_TO_USINT(X);
    	(* calculate the value of the digit *)
    	IF intX > 47 AND intX < 58 THEN
    		HEX_TO_BYTE := USINT_TO_BYTE(BYTE_TO_USINT(SHL(HEX_TO_BYTE,4)) + intX - 48);
    	ELSIF intX > 64 AND intX < 71 THEN
    		HEX_TO_BYTE := USINT_TO_BYTE(BYTE_TO_USINT(SHL(HEX_TO_BYTE,4)) + intX - 55);
    	ELSIF intX > 96 AND intX < 103 THEN
    		HEX_TO_BYTE := USINT_TO_BYTE(BYTE_TO_USINT(SHL(HEX_TO_BYTE,4)) + intX - 87);
    	END_IF
    	pt ACCESS (ADR(pt) + 1);
    END_FOR

    (* revision histroy
    hm	18. jun. 2008	rev 1.0
    	original release

    hm	20. sep.2008	rev 1.1
    	changed length of input string from 20 to 5

    *)

END_FUNCTION

(* ---- HEX_TO_DWORD.st ---- *)
FUNCTION HEX_TO_DWORD
    (*http://www.oscat.de/images/OSCATBasic/oscat_basic333_en.pdf#page=165*)
    pt ACCESS ADR(HEX);
    stop := LEN(HEX);
    FOR i := 1 TO stop DO
    	(* read the first character and subtract 48 to get value in decimal 0 = 48 *)
    	X := pt;
        intX := BYTE_TO_USINT(X);
    	(* calculate the value of the digit *)
    	IF intX > 47 AND intX < 58 THEN
    		HEX_TO_DWORD := UDINT_TO_DWORD(DWORD_TO_UDINT(SHL(HEX_TO_DWORD,4)) + intX - 48);
    	ELSIF intX > 64 AND intX < 71 THEN
    		HEX_TO_DWORD := UDINT_TO_DWORD(DWORD_TO_UDINT(SHL(HEX_TO_DWORD,4)) + intX - 55);
    	ELSIF intX > 96 AND intX < 103 THEN
    		HEX_TO_DWORD := UDINT_TO_DWORD(DWORD_TO_UDINT(SHL(HEX_TO_DWORD,4)) + intX - 87);
    	END_IF
    	pt ACCESS (ADR(pt) + 1);
    END_FOR

    (* revision histroy
    hm	2.10.2007		rev 1.0
    	original release

    hm	19.11.2007		rev 1.1
    	changed type of function from int to dword

    hm 	4. mar 2008		rev 1.2
    	added support for a..f and return 0 for invalid string

    hm	29. mar. 2008	rev 1.3
    	changed STRING to STRING(8)

    hm	18. jun. 2008	rev 1.4
    	changed input HEX to STRING(20)
    	function now ignores wrong characters
    *)

END_FUNCTION

(* ---- HOUR.st ---- *)
FUNCTION HOUR
    (*http://www.oscat.de/images/OSCATBasic/oscat_basic333_en.pdf#page=124*)
    HOUR := UDINT_TO_INT(TOD_TO_UDINT(ITOD) / 3600000);

    (* change history
    hm 4. aug 2006	rev 1.0
    	original version

    hm 2.10.2006 	rev 1.1
    	changed name of input to ITOD

    *)
END_FUNCTION

(* ---- HOUR_OF_DT.st ---- *)
FUNCTION HOUR_OF_DT
    (*http://www.oscat.de/images/OSCATBasic/oscat_basic333_en.pdf#page=125*)
    HOUR_OF_DT := UDINT_TO_INT((DT_TO_UDINT(XDT) MOD 86400) / 3600);

    (* revision history
    hm		6.9.2008	rev 1.0
    	original version

    *)
END_FUNCTION

(* ---- HOUR_TO_TIME.st ---- *)
FUNCTION HOUR_TO_TIME
    (*http://www.oscat.de/images/OSCATBasic/oscat_basic333_en.pdf#page=125*)
    HOUR_TO_TIME := DWORD_TO_TIME(REAL_TO_DWORD(IN * 3600000));

    (* revision history
    hm		4. aug 2006	rev 1.0
    	original version

    hm	14. mar. 2008	rev 1.1
    	rounded the input after the last digit

    hm	24. feb. 2009	rev 1.2
    	changed input to IN
    *)
END_FUNCTION

(* ---- HOUR_TO_TOD.st ---- *)
FUNCTION HOUR_TO_TOD
    (*http://www.oscat.de/images/OSCATBasic/oscat_basic333_en.pdf#page=125*)
    HOUR_TO_TOD := DWORD_TO_TOD(REAL_TO_DWORD(IN * 3600000));

    (* revision history
    hm	4. aug. 2006	rev 1.0
    	original version

    hm	14. mar. 2008	rev 1.1
    	rounded the input after the last digit

    hm	24. feb. 2009	rev 1.2
    	changed input to IN
    *)
END_FUNCTION

(* ---- HYPOT.st ---- *)
FUNCTION HYPOT
    (*http://www.oscat.de/images/OSCATBasic/oscat_basic333_en.pdf#page=55*)
    HYPOT := SQRT(X*X + Y*Y);

    (* revision history
    hm	21. feb 2008	rev 1.0
    	original version

    *)

END_FUNCTION

(* ---- INC.st ---- *)
FUNCTION INC
    (*http://www.oscat.de/images/OSCATBasic/oscat_basic333_en.pdf#page=55*)
    INC := (X + D + M + 1) MOD (M + 1);

    (* revision history
    hm	7. feb 2007		REV 1.0
    	original version

    hm	15. jan 2008	rev 1.1
    	allow for neagtive increment

    *)
END_FUNCTION

(* ---- INC1.st ---- *)
FUNCTION INC1
    (*http://www.oscat.de/images/OSCATBasic/oscat_basic333_en.pdf#page=56*)
    IF X >= N - 1 THEN
    	INC1 := 0;
    ELSE
    	INC1 := X + 1;
    END_IF

    (* revision history
    hm	13. oct. 2008	rev 1.0
    	original version

    hm	22. oct. 2008	rev 1.1
    	added statement to return value for compatibility reasons

    hm	23. feb. 2009	rev 1.2
     	when INC1 is called with X >= N inc will continue with 0
    *)
END_FUNCTION

(* ---- INC2.st ---- *)
FUNCTION INC2
    (*http://www.oscat.de/images/OSCATBasic/oscat_basic333_en.pdf#page=56*)
    tmp := U - L + 1;
    INC2 := (X + D - L + tmp) MOD tmp + L;

    (* revision history
    hm	29. jun. 2008		REV 1.0
    	original version

    *)
END_FUNCTION

(* ---- INT_TO_BCDC.st ---- *)
FUNCTION INT_TO_BCDC
    (*http://www.oscat.de/images/OSCATBasic/oscat_basic333_en.pdf#page=227*)
    INT_TO_BCDC := SHL(INT_TO_BYTE(IN / INT#10),4) OR INT_TO_BYTE(IN MOD INT#10);

    (* revision history
    hm	13.12.2007
    	original version

    hm	30.6.2008	rev 1.1
    	changed name INT_TO_BCD to INT_TO_BCDC to avoid collision with util.lib
    	corrected error IN code

    *)
END_FUNCTION

(* ---- INV.st ---- *)
FUNCTION INV
    (*http://www.oscat.de/images/OSCATBasic/oscat_basic333_en.pdf#page=57*)
    IF X <> 0.0 THEN INV := 1.0 / X; END_IF

    (* revision history
    hm	26. oct. 2008	rev 1.0
    	original version

    hm	10. mar. 2009	rev 1.1
    	real constants updated to new systax using dot

    *)

END_FUNCTION

(* ---- IS_ALNUM.st ---- *)
FUNCTION IS_ALNUM
    (*http://www.oscat.de/images/OSCATBasic/oscat_basic333_en.pdf#page=165*)
    pt ACCESS ADR(STR);
    L := LEN(STR);
    FOR pos := 1 TO L DO
    	IF NOT (ISC_ALPHA(pt) OR ISC_NUM(pt)) THEN
    		IS_ALNUM := FALSE;
    		RETURN;
    	END_IF
        	pt ACCESS (ADR(pt) + 1);
    END_FOR
    IS_ALNUM := L > 0;

    (* revision history
    hm	29. feb 2008	rev 1.0
    	original version

    hm	29. mar. 2008	rev 1.1
    	changed STRING to STRING(STRING_LENGTH)
    *)
END_FUNCTION

(* ---- IS_ALPHA.st ---- *)
FUNCTION IS_ALPHA
    (*http://www.oscat.de/images/OSCATBasic/oscat_basic333_en.pdf#page=165*)
    pt ACCESS ADR(STR);
    L := LEN(STR);
    FOR pos := 1 TO L DO
    	IF NOT ISC_ALPHA(pt) THEN
    		IS_ALPHA := FALSE;
    		RETURN;
    	END_IF
        pt ACCESS (ADR(pt) + 1);
    END_FOR
    IS_ALPHA := L > 0;

    (* revision history
    hm	29. feb 2008	rev 1.0
    	original version

    hm	29. mar. 2008	rev 1.1
    	changed STRING to STRING(STRING_LENGTH)
    *)
END_FUNCTION

(* ---- IS_CC.st ---- *)
FUNCTION IS_CC
    (*http://www.oscat.de/images/OSCATBasic/oscat_basic333_en.pdf#page=166*)
    L := LEN(STR);
    FOR pos := 1 TO L DO
    	IF FIND(CMP,MID(STR,1,pos)) = 0 THEN RETURN; END_IF
    END_FOR
    IS_CC := L > 0;

    (* revision history
    hm	19. mar 2008	rev 1.0
    	original version

    hm	29. mar. 2008	rev 1.1
    	changed STRING to STRING(STRING_LENGTH)
    *)
END_FUNCTION

(* ---- IS_CTRL.st ---- *)
FUNCTION IS_CTRL
    (*http://www.oscat.de/images/OSCATBasic/oscat_basic333_en.pdf#page=166*)
    pt ACCESS ADR(STR);
    L := LEN(STR);
    FOR pos := 1 TO L DO
    	IF NOT ISC_CTRL(pt) THEN
    		IS_CTRL := FALSE;
    		RETURN;
    	END_IF
        pt ACCESS (ADR(pt) + 1);
    END_FOR
    IS_CTRL := L > 0;

    (* revision history
    hm	29. feb. 2008	rev 1.0
    	original version

    hm	29. mar. 2008	rev 1.1
    	changed STRING to STRING(STRING_LENGTH)
    *)
END_FUNCTION

(* ---- IS_HEX.st ---- *)
FUNCTION IS_HEX
    (*http://www.oscat.de/images/OSCATBasic/oscat_basic333_en.pdf#page=167*)
    pt ACCESS ADR(STR);
    L := LEN(STR);
    FOR pos := 1 TO L DO
    	IF NOT ISC_HEX(pt) THEN
    		IS_HEX := FALSE;
    		RETURN;
    	END_IF
        	pt ACCESS (ADR(pt) + 1);
    END_FOR
    IS_HEX := L > 0;

    (* revision history
    hm	29. feb 2008	rev 1.0
    	original version

    hm	29. mar. 2008	rev 1.1
    	changed STRING to STRING(STRING_LENGTH)
    *)
END_FUNCTION

(* ---- IS_LOWER.st ---- *)
FUNCTION IS_LOWER
    (*http://www.oscat.de/images/OSCATBasic/oscat_basic333_en.pdf#page=167*)
    pt ACCESS ADR(STR);
    l := LEN(STR);
    FOR pos := 1 TO l DO
    	IF NOT ISC_LOWER(pt) THEN
    		IS_LOWER := FALSE;
    		RETURN;
    	END_IF
        	pt ACCESS (ADR(pt) + 1);
    END_FOR
    IS_LOWER := l > 0;

    (* revision history
    hm	29. feb 2008	rev 1.0
    	original version

    hm	29. mar. 2008	rev 1.1
    	changed STRING to STRING(STRING_LENGTH)
    *)
END_FUNCTION

(* ---- IS_NCC.st ---- *)
FUNCTION IS_NCC
    (*http://www.oscat.de/images/OSCATBasic/oscat_basic333_en.pdf#page=168*)
    L := LEN(STR);
    FOR pos := 1 TO L DO
    	IF FIND(CMP,MID(STR,1,pos)) > 0 THEN RETURN; END_IF
    END_FOR
    IS_NCC := TRUE;

    (* revision history
    hm	19. mar 2008	rev 1.0
    	original version

    hm	29. mar. 2008	rev 1.1
    	changed STRING to STRING(STRING_LENGTH)
    *)
END_FUNCTION

(* ---- IS_NUM.st ---- *)
FUNCTION IS_NUM
    (*http://www.oscat.de/images/OSCATBasic/oscat_basic333_en.pdf#page=168*)
    pt ACCESS ADR(STR);
    L := LEN(STR);
    FOR pos := 1 TO L DO
    	IF NOT ISC_NUM(pt) THEN
    		IS_NUM := FALSE;
    		RETURN;
    	END_IF
        	pt ACCESS (ADR(pt) + 1);
    END_FOR
    IS_NUM := L > 0;

    (* revision history
    hm	29. feb 2008	rev 1.0
    	original version

    hm	29. mar. 2008	rev 1.1
    	changed STRING to STRING(STRING_LENGTH)
    *)
END_FUNCTION

(* ---- IS_SORTED.st ---- *)
FUNCTION IS_SORTED
    (*http://www.oscat.de/images/OSCATBasic/oscat_basic333_en.pdf#page=82*)
    stop := UINT_TO_INT(SHR(SIZE,2)-2);
    FOR i := 0 TO stop DO
    	IF PT[i] > PT[i+1] THEN
    		IS_SORTED := FALSE;
    		RETURN;
    	END_IF
    END_FOR

    IS_SORTED := TRUE;

    (* revision history

    hm 	29. mar. 2008 	rev 1.0
    	original version

    hm	4. apr. 2008	rev 1.1
    	added type conversion to avoid warnings under codesys 3.0
    *)

END_FUNCTION

(* ---- IS_UPPER.st ---- *)
FUNCTION IS_UPPER
    (*http://www.oscat.de/images/OSCATBasic/oscat_basic333_en.pdf#page=169*)
    pt ACCESS ADR(STR);
    L := LEN(STR);
    FOR pos := 1 TO L DO
    	IF NOT ISC_UPPER(pt) THEN
    		IS_UPPER := FALSE;
    		RETURN;
    	END_IF
        pt ACCESS (ADR(pt) + 1);
    END_FOR
    IS_UPPER := L > 0;

    (* revision history
    hm	29. feb 2008	rev 1.0
    	original version

    hm	29. mar. 2008	rev 1.1
    	changed STRING to STRING(STRING_LENGTH)
    *)
END_FUNCTION

(* ---- ISC_ALPHA.st ---- *)
FUNCTION ISC_ALPHA
    (*http://www.oscat.de/images/OSCATBasic/oscat_basic333_en.pdf#page=169*)
    IF cEXTENDED_ASCII THEN
    	ISC_ALPHA := (IN > 64 AND IN < 91) OR (IN > 191  AND IN <> 215 AND IN <> 247) OR (IN > 96 AND IN < 123);
    ELSE
    	ISC_ALPHA := (IN > 64 AND IN < 91) OR (IN > 96 AND IN < 123);
    END_IF

    (* revision history
    hm	6. mar. 2008	rev 1.0
    	original version

    hm	19. oct. 2008	rev 1.1
    	changes setup constants
    *)

END_FUNCTION

(* ---- ISC_CTRL.st ---- *)
FUNCTION ISC_CTRL
    (*http://www.oscat.de/images/OSCATBasic/oscat_basic333_en.pdf#page=170*)
    ISC_CTRL := IN < 32 OR IN = 127;

    (* revision history
    hm		6. mar. 2008	rev 1.0
    	original version

    *)
END_FUNCTION

(* ---- ISC_HEX.st ---- *)
FUNCTION ISC_HEX
    (*http://www.oscat.de/images/OSCATBasic/oscat_basic333_en.pdf#page=170*)
    ISC_HEX := (IN > 47 AND IN < 58) OR (IN > 64 AND IN < 71) OR (IN > 96 AND IN < 103);

    (* revision history
    hm		6. mar. 2008	rev 1.0
    	original version

    *)
END_FUNCTION

(* ---- ISC_LOWER.st ---- *)
FUNCTION ISC_LOWER
    (*http://www.oscat.de/images/OSCATBasic/oscat_basic333_en.pdf#page=171*)
    IF cEXTENDED_ASCII THEN
    	ISC_LOWER := ((IN > 96) AND (IN < 123)) OR ((IN > 222) AND (IN <> 247));
    ELSE
    	ISC_LOWER := ((IN > 96) AND (IN < 123));
    END_IF

    (* revision history
    hm	6. mar. 2008	rev 1.0
    	original version

    hm	19. oct. 2008	rev 1.1
    	changes setup constants
    *)
END_FUNCTION

(* ---- ISC_NUM.st ---- *)
FUNCTION ISC_NUM
    (*http://www.oscat.de/images/OSCATBasic/oscat_basic333_en.pdf#page=171*)
    ISC_NUM := IN > 47 AND IN < 58;

    (* revision history
    hm		6. mar. 2008	rev 1.0
    	original version

    *)
END_FUNCTION

(* ---- ISC_UPPER.st ---- *)
FUNCTION ISC_UPPER
    (*http://www.oscat.de/images/OSCATBasic/oscat_basic333_en.pdf#page=172*)
    IF cEXTENDED_ASCII THEN
    	ISC_UPPER :=  ((IN > 64) AND (IN < 91)) OR (((IN > 191) AND (IN < 223)) AND (IN <> 215));
    ELSE
    	ISC_UPPER := ((IN > 64) AND (IN < 91));
    END_IF

    (* revision history
    hm	6. mar. 2008	rev 1.0
    	original version

    hm	19. oct. 2008	rev 1.1
    	changes setup constants

    *)
END_FUNCTION

(* ---- JD2000.st ---- *)
FUNCTION JD2000
    (*http://www.oscat.de/images/OSCATBasic/oscat_basic333_en.pdf#page=126*)
    JD2000 := UDINT_TO_REAL(DT_TO_UDINT(DTI) - 946728000) / 86400.0;

    (* revision histroy
    hm	15. jul. 2008	rev 1.0
    	original release

    *)

END_FUNCTION

(* ---- K_TO_C.st ---- *)
FUNCTION K_TO_C
    (*http://www.oscat.de/images/OSCATBasic/oscat_basic333_en.pdf#page=366*)
    K_TO_C := KELVIN + cT0;

    (* revision history

    hm	4. aug 2006	rev 1.0
    	original version

    hm	19. aug 2009	rev 1.1
    	fixed calculation error

    *)

END_FUNCTION

(* ---- KMH_TO_MS.st ---- *)
FUNCTION KMH_TO_MS
    (*http://www.oscat.de/images/OSCATBasic/oscat_basic333_en.pdf#page=366*)
    KMH_TO_MS := KMH * 0.2777777777777;

    (* revision history
    hm	4. feb 2007		rev 1.0
    	original version

    hm	6. jan 2008		rev 1.1
    	improved performance

    *)

END_FUNCTION

(* ---- LAMBERT_W.st ---- *)
FUNCTION LAMBERT_W
    (*http://www.oscat.de/images/OSCATBasic/oscat_basic333_en.pdf#page=58*)
    (* check for valid input and return -1000 if too low *)
    IF X < -0.367879441171442 THEN
    	LAMBERT_W := -1000.0;
    	RETURN;
    (* return 0 if X = 0 *)
    ELSIF X = 0.0 THEN
    	RETURN;
    (* first an estimate is calculated *)
    ELSIF X <= 500.0 THEN
    	w := LN(X + 1.0);
    	w := 0.665 * (1.0 + 0.0195 * w) * w + 0.04;
    ELSE
    	w := LN(X - 4.0) - (1.0 - 1.0/LN(X)) * LN(LN(X));
    END_IF
    (* use estimate to calculate exact result *)
    FOR i := 0 TO 5 DO
    	ewx := EXP(w);
    	we := w * ewx - X;
    	w1e := (w+1.0) * ewx;
    	last := REAL_TO_DW(w) AND 16#FFFF_FFFC;
    	w := w - (we / (w1e - (w+2.0) * we / (2.0 * w + 2.0)));
    	IF (REAL_TO_DW(w) AND 16#FFFF_FFFC) = last THEN EXIT; END_IF
    END_FOR
    LAMBERT_W := w;

    (* revision hisdtory
    hm	26. oct. 2008	rev 1.0
    	original version

    hm	10. mar. 2009	rev 1.1
    	real constants updated to new systax using dot

    *)
END_FUNCTION

(* ---- LANGEVIN.st ---- *)
FUNCTION LANGEVIN
    (*http://www.oscat.de/images/OSCATBasic/oscat_basic333_en.pdf#page=58*)
    IF X = 0.0 THEN
    	LANGEVIN := 0.0;
    ELSE
    	LANGEVIN := COTH(X) - 1.0 / X;
    END_IF

    (* revision history
    hm	10.12.2007	rev 1.0
    	original version

    hm	11. mar 2008	rev 1.1
    	changed formula to avoid problems when X = 0

    hm	10. mar. 2009	rev 1.2
    	real constants updated to new systax using dot

    *)
END_FUNCTION

(* ---- LEAP_DAY.st ---- *)
FUNCTION LEAP_DAY
    (*http://www.oscat.de/images/OSCATBasic/oscat_basic333_en.pdf#page=126*)
    LEAP_DAY := DATE_TO_UDINT(IDATE) MOD 126230400 = 68169600;

    (* change history

    hm 	15. jun. 2008	rev 1.0
    	original version

    hm	7. oct. 2008	rev 1.1
    	changed function month to month_of_date

    hm	24. jan. 2011	rev 1.2
    	improved performance
    *)
END_FUNCTION

(* ---- LEAP_OF_DATE.st ---- *)
FUNCTION LEAP_OF_DATE
    (*http://www.oscat.de/images/OSCATBasic/oscat_basic333_en.pdf#page=127*)
    LEAP_OF_DATE := SHL(((DATE_TO_UDINT(IDATE) + 43200) / 31557600), 30) = 16#80000000;

    (* change history

    2.10.2006		rev 1.1
    the function now calls leap_year to accomodate further accuracy.
    the function now works for any year from 1970 to 2100

    8. jan 2008		rev 1.2
    	improved code for better performance

    28. jan. 2011	rev 1.3
    	improved performance
    *)
END_FUNCTION

(* ---- LEAP_YEAR.st ---- *)
FUNCTION LEAP_YEAR
    (*http://www.oscat.de/images/OSCATBasic/oscat_basic333_en.pdf#page=127*)
    LEAP_YEAR := SHL(YR,14) = 0;

    (* this code was used prior to rev 1.1

    IF YR MOD 400 = 0 THEN LEAP_YEAR := TRUE;
    ELSIF YR MOD 100 = 0 THEN LEAP_YEAR := FALSE;
    ELSIF YR MOD 4 =0 THEN LEAP_YEAR := TRUE;
    ELSE LEAP_YEAR := FALSE;
    END_IF

    *)

    (* change history

    hm 	2.10.2006		rev 1.1
    	the function now works for any year from 1970 up to 2100

    hm	1. oct 2007		rev 1.2
    	chaged code for higher performance
    *)
END_FUNCTION

(* ---- LINEAR_INT.st ---- *)
FUNCTION LINEAR_INT
    (*http://www.oscat.de/images/OSCATBasic/oscat_basic333_en.pdf#page=101*)
    (*make sure n is bound within the array size *)
    PTS := MIN(PTS,20);

    (* calculate the linear segement interpolation *)
    i := 2;
    (* search for segment and calculate output
    	below and above the defined segments we interpolate the last segment *)
    WHILE (i < PTS) AND (XY[i,0] < X) DO
    	i := i + 1;
    END_WHILE

    (* calculate the output value on the corresponding segment coordinates *)
    LINEAR_INT := ((XY[i,1] - XY[i-1,1]) * X - XY[i,1] * XY[i-1,0] + XY[i-1,1] * XY[i,0]) / (XY[i,0] - XY[i-1,0]);

    (* revision history
    hm	7. oct 2007		rev 1.0
    	original version

    hm	27 dec 2007		rev 1.1
    	changed code for better performance
    *)

END_FUNCTION

(* ---- LIST_CLEAN.st ---- *)
FUNCTION LIST_CLEAN
    (*http://www.oscat.de/images/OSCATBasic/oscat_basic333_en.pdf#page=485*)
    pt ACCESS ADR(LIST);

    FOR read := 1 TO LIST_LENGTH DO
    	c := pt[read];								(* read character from LIST *)
    	IF c = 0 THEN EXIT;						(* exit the loop if character definbes end of string *)
    	ELSIF c <> SEP OR SEP <> last THEN	(* copy element from read to write position unless a double SEP character is present *)
    		pt[write] := c;
    		write := write + 1;
    	END_IF
    	last := c;									(* remember last character *)
    END_FOR

    IF last = SEP THEN write := write - 1; END_IF		(* if last character is SEP then delete empty element at end *)
    IF write <= STRING_LENGTH THEN pt[write] := 0;	 END_IF		(* terminate string with 0 *)

    LIST_CLEAN := TRUE;						(* retrun TRUE *)

    (* revision histroy
    hm	28. jun. 2008	rev 1.0
    	original release

    hm	19. jan. 2011	rev 1.1
    	changed string(255) to string(LIST_LENGTH)

    hm	21. mar. 2011	rev 2.0
    	all elements start with SEP

    *)

END_FUNCTION

(* ---- LIST_GET.st ---- *)
FUNCTION LIST_GET
    (*http://www.oscat.de/images/OSCATBasic/oscat_basic333_en.pdf#page=485*)
    pt ACCESS ADR(LIST);							(* load pointers *)
    po ACCESS ADR(LIST_GET);

    REPEAT
    	c := pt[i];
    	IF cnt = POS THEN						(* copy element to output string *)
    		IF c = SEP  THEN EXIT; END_IF		(* next element stop copy and finish *)
    		po[o] := c;
    		o := o + 1;
    	ELSIF c = SEP THEN
    		cnt := cnt + 1;
    	END_IF
    	i := i + 1;
    UNTIL
    	(i = LIST_LENGTH) OR (c = 0)
    END_REPEAT
    po[o] := 0;						(* close the output string *)

    (* revision histroy
    hm	20. jun. 2008	rev 1.0
    	original release

    hm	19. jan. 2011	rev 1.1
    	changed string(255) to strring(LIST_LENGTH)

    hm	21. mar. 2011	rev 2.0
    	all LIST elements start with SEP
    *)

END_FUNCTION

(* ---- LIST_INSERT.st ---- *)
FUNCTION LIST_INSERT
    (*http://www.oscat.de/images/OSCATBasic/oscat_basic333_en.pdf#page=486*)
    (* load pointers *)
    pt ACCESS ADR(LIST);

    IF LEN(INS) + 1 + LEN(LIST) > LIST_LENGTH THEN
    	LIST_INSERT := FALSE;
    ELSE
    	LIST_INSERT := TRUE;
    	(* search for position *)
    	WHILE read < LIST_LENGTH DO
    		IF cnt >= POS THEN
    			CHR_TO_STRING(SEP, sx);
    			INS := CONCAT(sx, INS);
    			LIST := INSERT(LIST, INS, read - 1);
    			LIST_INSERT := TRUE;
    			RETURN;
    		END_IF
    		IF pt[read]  = 0 THEN				(* LIST is too short add empty element *)
    			pt[read] := SEP;
    			pt[read + 1] := 0;
    		END_IF
    		read := read + 1;
    		IF pt[read] = SEP OR pt[read] = 0 THEN cnt := cnt + 1; END_IF
    	END_WHILE
    END_IF

    (* revision histroy
    hm	28. jun. 2008	rev 1.0
    	original release

    hm	17. dec. 2008	rev 1.1
    	changes name of function chr to chr_to_string

    hm	19. jan. 2011	rev 1.2
    	changed string(255) to string(LIST_LENGTH)

    hm	21. mar. 2011	rev 2.0
    	all LIST elements start with SEP

    *)

END_FUNCTION

(* ---- LIST_LEN.st ---- *)
FUNCTION LIST_LEN
    (*http://www.oscat.de/images/OSCATBasic/oscat_basic333_en.pdf#page=487*)
    pt ACCESS ADR(LIST);
    LIST_LEN := 0;
    REPEAT
    	c := pt[pos];
    	IF c = SEP THEN LIST_LEN := LIST_LEN + 1; END_IF
    	pos := pos + 1;
    UNTIL
    	c = 0 OR pos > LIST_LENGTH
    END_REPEAT

    (* revision histroy
    hm	25. jun. 2008	rev 1.0
    	original release

    hm	16. oct. 2008	rev 1.1
    	fixed a problem where LIST_LEN would only work up to LIST_LENGTH

    hm	19. jan. 2001	rev 1.2
    	changed string(255) to string(LIST_LENGTH)

    hm	21. mar. 2011	rev 2.0
    	all LIST elements start with SEP

    *)

END_FUNCTION

(* ---- LIST_RETRIEVE.st ---- *)
FUNCTION LIST_RETRIEVE
    (*http://www.oscat.de/images/OSCATBasic/oscat_basic333_en.pdf#page=488*)
    (* load pointers *)
    pt ACCESS ADR(LIST);
    po ACCESS ADR(RETVAL);

    IF POS > 0 THEN
    	FOR i := 1 TO LIST_LENGTH DO
    		c := pt[i];
    		IF c = 0 THEN
    			po[o] := 0;
    			IF cnt < POS THEN pt[w + 1] := 0; ELSE pt[w] := 0; END_IF
                LIST_RETRIEVE := TRUE;
    			RETURN;
    		ELSIF cnt = POS AND c <> SEP THEN				(* we have found the element *)
    			po[o] := pt[i];
    			o := o + 1;
    		ELSIF cnt >= POS THEN
    			pt[w] := c;
    			w := w + 1;
    		ELSE
    			w := i;
    		END_IF
    		IF c = SEP THEN cnt := cnt + 1; END_IF
    	END_FOR
    ELSE
    	RETVAL := '';
        LIST_RETRIEVE := FALSE;
    END_IF

    (* revision histroy
    hm	28. jun. 2008	rev 1.0
    	original release

    hm	19. jan. 2011	rev 1.1
    	changed string(255) to string(LIST_LENGTH)

    hm	21. mar. 2011	rev 2.0
    	all elements start with SEP
    *)

END_FUNCTION

(* ---- LOWERCASE.st ---- *)
FUNCTION LOWERCASE
    (*http://www.oscat.de/images/OSCATBasic/oscat_basic333_en.pdf#page=172*)
    PT ACCESS ADR(RETVAL);
    RETVAL := STR;
    l := LEN(STR);
    FOR pos := 1 TO l DO
    	PT := TO_LOWER(PT);
    	PT ACCESS (ADR(PT) + 1);
    END_FOR
    LOWERCASE := TRUE;

    (* revision histroy
    hm	6. oct. 2006	rev 1.0
    	original release

    hm	4. feb. 2008	rev 1.1
    	improved performance
    	added Ä.Ö,Ü

    hm	6. mar. 2008	rev 1.2
    	added support for exteded Ascii

    hm	29. mar. 2008	rev 1.3
    	changed STRING to STRING(STRING_LENGTH)
    *)

END_FUNCTION

(* ---- LTIME_TO_UTC.st ---- *)
FUNCTION LTIME_TO_UTC
    (*http://www.oscat.de/images/OSCATBasic/oscat_basic333_en.pdf#page=128*)
    LTIME_TO_UTC := UDINT_TO_DT(DT_TO_UDINT(LOCAL_TIME) - INT_TO_UDINT(TIME_ZONE_OFFSET) * 60);
    IF DST THEN LTIME_TO_UTC := LTIME_TO_UTC - T#1h; END_IF

    (* revision history
    hm 5.7.2007		rev 1.0
    	original version

    hm 5.11.2007		rev 1.1
    	replaced literal constant with variable because of error in möller ecp4 compiler

    hm	12.nov 2007	rev 1.2
    	changed Type of TIME_ZONE_OFFSET from time to int to allow for time zones with negative offset

    hm	8. dec 2007	rev 1.3
    	corrected a problem with TIME_ZONE_OFFSET

    hm	14. oct. 2008	rev 1.4
    	changed TIME_ZONE_OFFSET from int to real to allow for half hour offset

    hm	20. oct. 2006	rev 1.5
    	changed TIME_ZONE_OFFSET from Real to INT, now in Minutes

    hm	27. feb. 2009	rev 1.6
    	added type conversions to avoid warnings under codesys 3.0

    ks	13. nov. 2009	rev 1.7
    	corrected error in formula

    *)
END_FUNCTION

(* ---- MANUAL.st ---- *)
FUNCTION MANUAL
    (*http://www.oscat.de/images/OSCATBasic/oscat_basic333_en.pdf#page=463*)
    MANUAL := NOT OFF AND (IN OR ON);

    (* revision history
    hm	21. nov 2008	rev 1.0
    	original version

    *)
END_FUNCTION

(* ---- MAX3.st ---- *)
FUNCTION MAX3
    (*http://www.oscat.de/images/OSCATBasic/oscat_basic333_en.pdf#page=59*)
    MAX3 := MAX(MAX(IN1,IN2),IN3);

    (* revision history
    hm	1.1.2007	rev 1.0
    	original release

    hm	18. mar. 2011	rev 1.1
    	improve performance

    *)
END_FUNCTION

(* ---- MID3.st ---- *)
FUNCTION MID3
    (*http://www.oscat.de/images/OSCATBasic/oscat_basic333_en.pdf#page=59*)
    IF IN1 > IN2 THEN MID3 := IN1; IN1 := IN2; IN2 := MID3; END_IF
    IF IN2 > IN3 THEN IN2 := IN3; END_IF
    MID3 := SEL(IN1 > IN2, IN2, IN1);

    (*
    hm	1.1.2007	rev 1.1
    	rewrote the function for better performance

    hm	18. mar. 2011	rev 1.2
    	improve performance
    *)
END_FUNCTION

(* ---- MIN3.st ---- *)
FUNCTION MIN3
    (*http://www.oscat.de/images/OSCATBasic/oscat_basic333_en.pdf#page=60*)
    MIN3 := MIN(MIN(IN1,IN2),IN3);

    (* revision history
    hm	1.1.2007	rev 1.0
    	original release

    hm	18. mar. 2011	rev 1.1
    	improve performance

    *)
END_FUNCTION

(* ---- MINUTE.st ---- *)
FUNCTION MINUTE
    (*http://www.oscat.de/images/OSCATBasic/oscat_basic333_en.pdf#page=128*)
    MINUTE := UDINT_TO_INT(TOD_TO_UDINT(ITOD) / 60000 - TOD_TO_UDINT(ITOD) / 3600000 * 60);

    (* change history

    2.10.2006 changes name of input to ITOD

    *)
END_FUNCTION

(* ---- MINUTE_OF_DT.st ---- *)
FUNCTION MINUTE_OF_DT
    (*http://www.oscat.de/images/OSCATBasic/oscat_basic333_en.pdf#page=128*)
    MINUTE_OF_DT := UDINT_TO_INT(DT_TO_UDINT(XDT) MOD 3600) / 60;

    (* revision history
    hm		6.9.2008	rev 1.0
    	original version

    *)
END_FUNCTION

(* ---- MINUTE_TO_TIME.st ---- *)
FUNCTION MINUTE_TO_TIME
    (*http://www.oscat.de/images/OSCATBasic/oscat_basic333_en.pdf#page=129*)
    MINUTE_TO_TIME := DWORD_TO_TIME(REAL_TO_DWORD(IN * 60000.0));

    (* revision history
    hm	4. aug 2006	rev 1.0
    	original version

    hm	14. mar 2008	rev 1.1
    	rounded the input after the last digit

    hm	24. feb. 2009	rev 1.2
    	changed input to IN

    *)
END_FUNCTION

(* ---- MIRROR.st ---- *)
FUNCTION MIRROR
    (*http://www.oscat.de/images/OSCATBasic/oscat_basic333_en.pdf#page=174*)
    pi ACCESS ADR(STR);
    po ACCESS ADR(RETVAL);
    lx := LEN(STR);
    FOR i := lx TO 1 BY - 1 DO
    	po := pi[i];
    	po ACCESS (ADR(po) + 1);
    END_FOR
    (* close output string *)
    po:= 0;
    MIRROR := TRUE;

    (* revision histroy
    hm	4. feb. 2008	rev 1.0
    	original release

    hm	29. mar. 2008	rev 1.1
    	changed STRING to STRING(STRING_LENGTH)
    *)

END_FUNCTION

(* ---- MIX.st ---- *)
FUNCTION MIX
    (*http://www.oscat.de/images/OSCATBasic/oscat_basic333_en.pdf#page=281*)
    MIX := (1.0 - M) * A + M * B;

    (* revision history
    hm	19. Nov 2007	rev 1.0
    	original version

    hm	10. mar 2009	rev 1.1
    	real constants updated to new systax using dot

    *)
END_FUNCTION

(* ---- MODR.st ---- *)
FUNCTION MODR
    (*http://www.oscat.de/images/OSCATBasic/oscat_basic333_en.pdf#page=60*)
    IF DIVI = 0.0 THEN
    	MODR := 0.0;
    ELSE
    	MODR := IN - DINT_TO_REAL(FLOOR2(IN / DIVI)) * DIVI;
    END_IF

    (* revision history

    hm	4. aug.2006		rev 1.0

    hm	28. jan.2007	rev 1.1
    	MODR(x,0) will deliver the result 0

    hm	21. mar 2008	rev 1.2
    	use D_trunc for compatibility reasons

    hm	4. apr. 2008	rev 1.3
    	added type conversion to avoid warnings under codesys 3.0

    hm	31. oct. 2008	rev 1.4
    	changed algorithm to the more common version using floor instead of TRUNC

    hm	10. mar. 2009	rev 1.5
    	real constants updated to new systax using dot

    *)
END_FUNCTION

(* ---- MONTH_BEGIN.st ---- *)
FUNCTION MONTH_BEGIN
    (*http://www.oscat.de/images/OSCATBasic/oscat_basic333_en.pdf#page=129*)
    MONTH_BEGIN := UDINT_TO_DATE(DATE_TO_UDINT(IDATE) - INT_TO_UDINT(DAY_OF_MONTH(IDATE) - 1) * 86400);

    (* revision history
    hm	15. jun. 2008	rev 1.0
    	original version

    *)
END_FUNCTION

(* ---- MONTH_END.st ---- *)
FUNCTION MONTH_END
    (*http://www.oscat.de/images/OSCATBasic/oscat_basic333_en.pdf#page=130*)
    MONTH_END := UDINT_TO_DATE(DATE_TO_UDINT(SET_DATE(YEAR_OF_DATE(IDATE),MONTH_OF_DATE(IDATE)+1,1)) - 86400);

    (* revision history
    hm	15. jun. 2008	rev 1.0
    	original version

    hm	7. oct. 2008	rev 1.1
    	changed function year to year_of_date
    	changed function month to month_of_date

    *)
END_FUNCTION

(* ---- MONTH_OF_DATE.st ---- *)
FUNCTION MONTH_OF_DATE
    (*http://www.oscat.de/images/OSCATBasic/oscat_basic333_en.pdf#page=130*)
    MONTH_OF_DATE := DAY_OF_YEAR(IDATE);
    IF MONTH_OF_DATE < 32 THEN
    	MONTH_OF_DATE := 1;
    ELSIF LEAP_OF_DATE(IDATE) THEN
    	MONTH_OF_DATE := (MONTH_OF_DATE * 53 + 1668) / 1623;
    ELSE
    	MONTH_OF_DATE := (MONTH_OF_DATE * 53 + 1700) / 1620;
    END_IF

    (* code for rev 1.2
    MONTH_OF_DATE := DAY_OF_YEAR(IDATE);
    IF LEAP_OF_DATE(IDATE) THEN
    	CASE MONTH_OF_DATE OF
    		1..31 	:	MONTH_OF_DATE := 1;
    		32..60	:	MONTH_OF_DATE := 2;
    		61..91	:	MONTH_OF_DATE := 3;
    		92..121 :	MONTH_OF_DATE := 4;
    		122..152:	MONTH_OF_DATE := 5;
    		153..182:	MONTH_OF_DATE := 6;
    		183..213:	MONTH_OF_DATE := 7;
    		214..244:	MONTH_OF_DATE := 8;
    		245..274:	MONTH_OF_DATE := 9;
    		275..305:	MONTH_OF_DATE := 10;
    		306..335:	MONTH_OF_DATE := 11;
    		336..366:	MONTH_OF_DATE := 12;
    	END_CASE
    ELSE
    	CASE MONTH_OF_DATE OF
    		1..31 	:	MONTH_OF_DATE := 1;
    		32..59	:	MONTH_OF_DATE := 2;
    		60..90	:	MONTH_OF_DATE := 3;
    		91..120 :	MONTH_OF_DATE := 4;
    		121..151:	MONTH_OF_DATE := 5;
    		152..181:	MONTH_OF_DATE := 6;
    		182..212:	MONTH_OF_DATE := 7;
    		213..243:	MONTH_OF_DATE := 8;
    		244..273:	MONTH_OF_DATE := 9;
    		274..304:	MONTH_OF_DATE := 10;
    		305..334:	MONTH_OF_DATE := 11;
    		335..365:	MONTH_OF_DATE := 12;
    	END_CASE
    END_IF
    *)

    (* revision history
    hm	1. aug 2006	rev 1.0
    	original version

    hm	1. okt 2007	rev 1.1
    	replaced old code (string conversion) with mathematics
    	the execution time is now multiple times faster.

    hm	7. oct. 2008	rev 1.2
    	changed name of function from month to MONTH_OF_DATE

    hm	27. mar. 2009	rev 1.3
    	new improved code

    *)
END_FUNCTION

(* ---- MONTH_TO_STRING.st ---- *)
FUNCTION MONTH_TO_STRING
    (*http://www.oscat.de/images/OSCATBasic/oscat_basic333_en.pdf#page=175*)
    IF LANG = 0 THEN ly := cLANGUAGE_DEFAULT; ELSE ly := MIN(LANG, cLANGUAGE_LMAX); END_IF
    IF MTH < 1 OR MTH > 12 THEN
    	RETURN;
    ELSIF LX = 0 THEN
    	RETVAL := cMONTHS[ly, MTH];
    ELSIF LX = 3 THEN
    	RETVAL := cMONTHS3[ly, MTH];
    END_IF
    MONTH_TO_STRING := TRUE;

    (* revisison history

    hm	21. sep. 2008	rev 1.0
    	original version

    hm	19. oct. 2008	rev 1.1
    	changed language setup constants
    *)
END_FUNCTION

(* ---- MS_TO_BFT.st ---- *)
FUNCTION MS_TO_BFT
    (*http://www.oscat.de/images/OSCATBasic/oscat_basic333_en.pdf#page=368*)
    MS_TO_BFT := REAL_TO_INT(EXPT(MS * 1.196172, 0.666667));

    (* revision history
    hm	12. 6. 2008		rev 1.0
    	original version

    *)
END_FUNCTION

(* ---- MS_TO_KMH.st ---- *)
FUNCTION MS_TO_KMH
    (*http://www.oscat.de/images/OSCATBasic/oscat_basic333_en.pdf#page=369*)
    MS_TO_KMH := MS * 3.6;

END_FUNCTION

(* ---- MUL_ADD.st ---- *)
FUNCTION MUL_ADD
    (*http://www.oscat.de/images/OSCATBasic/oscat_basic333_en.pdf#page=61*)
    MUL_ADD := X * K + O;

    (* revision history
    hm	28. feb 2007
    	original version

    hm	11.nov 2007		rev 1.1
    	deleted preset values for K and O this makes no sense for a function

    *)
END_FUNCTION

(* ---- MULTI_IN.st ---- *)
FUNCTION MULTI_IN
    (*http://www.oscat.de/images/OSCATBasic/oscat_basic333_en.pdf#page=317*)
    F1 :=  IN_1 > IN_MIN AND IN_1 < IN_MAX;
    F2 :=  IN_2 > IN_MIN AND IN_2 < IN_MAX;
    F3 :=  IN_3 > IN_MIN AND IN_3 < IN_MAX;

    CASE MODE OF
    0:	count := 0;
    	IF F1 THEN
    		count := count + 1;
    		MULTI_IN := IN_1;
    	ELSE
    		MULTI_IN := 0.0;
    	END_IF
    	IF F2 THEN
    		count := count + 1;
    		MULTI_IN := MULTI_IN + IN_2;
    	END_IF
    	IF F3 THEN
    		count := count + 1;
    		MULTI_IN := MULTI_IN + IN_3;
    	END_IF
    	MULTI_IN := SEL(count = 0, MULTI_IN / INT_TO_REAL(count), DEFAULT);

    1:	MULTI_IN := SEL(F1, DEFAULT, IN_1);

    2:	MULTI_IN := SEL(F2, DEFAULT, IN_2);

    3:	MULTI_IN := SEL(F3, DEFAULT, IN_3);

    4:	MULTI_IN := DEFAULT;

    5:	MULTI_IN := SEL(F1, IN_MAX, IN_1);
    	IF F2 AND IN_2 < MULTI_IN THEN MULTI_IN := IN_2; END_IF
    	IF F3 AND IN_3 < MULTI_IN THEN MULTI_IN := IN_3; END_IF
    	IF MULTI_IN = IN_MAX THEN MULTI_IN := DEFAULT; END_IF

    6:	MULTI_IN := SEL(F1, IN_MIN, IN_1);
    	IF F2 AND IN_2 > MULTI_IN THEN MULTI_IN := IN_2; END_IF
    	IF F3 AND IN_3 > MULTI_IN THEN MULTI_IN := IN_3; END_IF
    	IF MULTI_IN = IN_MIN THEN MULTI_IN := DEFAULT; END_IF

    7:	IF F1 AND F2 AND F3 THEN MULTI_IN := MID3(IN_1, IN_2, IN_3);
    	ELSIF F1 AND F2 THEN MULTI_IN := MIN(IN_1, IN_2);
    	ELSIF F1 AND F3 THEN MULTI_IN := MIN(IN_1, IN_3);
    	ELSIF F2 AND F3 THEN MULTI_IN := MIN(IN_2, IN_3);
    	ELSIF F1 THEN MULTI_IN := IN_1;
    	ELSIF F2 THEN MULTI_IN := IN_2;
    	ELSIF F3 THEN MULTI_IN := IN_3;
    	ELSE MULTI_IN := DEFAULT;
    	END_IF

    END_CASE

    (*
    hm 1.1.2007		rev 1.1
    	changed midr to mid3 function

    hm	14. 10. 2008	rev 1.2
    	corrected an error for IN_3 overrange detection
    	improved performance

    hm	11. mar. 2009	rev 1.3
    	changed real constants to use dot syntax

    hm	18. jul. 2009	rev 1.4
    	improved performance
    *)
END_FUNCTION

(* ---- MULTIME.st ---- *)
FUNCTION MULTIME
    (*http://www.oscat.de/images/OSCATBasic/oscat_basic333_en.pdf#page=130*)
    MULTIME := DWORD_TO_TIME(REAL_TO_DWORD(DWORD_TO_REAL(TIME_TO_DWORD(T))*M));

    (* revision history
    hm		2. oct 2006	rev 1.0
    	original version

    hm		14. mar 2008	rev 1.1
    	rounded the result after the last digit

    *)
END_FUNCTION

(* ---- MUX_2.st ---- *)
FUNCTION MUX_2
    (*http://www.oscat.de/images/OSCATBasic/oscat_basic333_en.pdf#page=229*)
    MUX_2 := SEL(A0, D0, D1);

    (*
    revision history:
    hm	5.10.2006		rev 1.1
    	changed to ST Langage for better portability.

    hm	16. oct. 2008	rev 1.2
    	improved performance

    *)
END_FUNCTION

(* ---- MUX_4.st ---- *)
FUNCTION MUX_4
    (*http://www.oscat.de/images/OSCATBasic/oscat_basic333_en.pdf#page=229*)
    IF A1 THEN
    	MUX_4 := SEL(A0, D2, D3);
    ELSE
    	MUX_4 := SEL(A0, D0, D1);
    END_IF

    (*
    revision history:
    hm 	5.10.2006		rev 1.1
    	rewritten to ST for better portability

    hm	16. oct. 2008	rev 1.2
    	improved performance

    *)
END_FUNCTION

(* ---- MUX_R2.st ---- *)
FUNCTION MUX_R2
    (*http://www.oscat.de/images/OSCATBasic/oscat_basic333_en.pdf#page=281*)
    MUX_R2 := SEL(A, IN0, IN1);

    (* revision history
    hm	19. jan. 2007	rev 1.0
    	original version

    hm	16. oct. 2008	rev 1.1
    	improved performance

    *)
END_FUNCTION

(* ---- MUX_R4.st ---- *)
FUNCTION MUX_R4
    (*http://www.oscat.de/images/OSCATBasic/oscat_basic333_en.pdf#page=282*)
    IF A1 THEN
    	MUX_R4 := SEL(A0, IN2, IN3);
    ELSE
    	MUX_R4 := SEL(A0, IN0, IN1);
    END_IF

    (* revision history
    hm	19. jan 2007	rev 1.0
    	original version

    hm	16. oct. 2008	rev 1.1
    	improved performance
    *)
END_FUNCTION

(* ---- NEGX.st ---- *)
FUNCTION NEGX
    (*http://www.oscat.de/images/OSCATBasic/oscat_basic333_en.pdf#page=61*)
    NEGX := -X;

    (* revision history
    hm	26. oct. 2008	rev 1.0
    	original version

    *)

END_FUNCTION

(* ---- OCT_TO_BYTE.st ---- *)
FUNCTION OCT_TO_BYTE
    (*http://www.oscat.de/images/OSCATBasic/oscat_basic333_en.pdf#page=175*)
    pt ACCESS ADR(OCT);
    stop := LEN(OCT);
    FOR i := 1 TO stop DO
    	(* read the first character and subtract 48 to get value in decimal 0 = 48 *)
    	X := pt;
        intX := BYTE_TO_USINT(X);
    	(* calculate the value of the digit *)
    	IF intX > 47 AND intX < 56 THEN
    		OCT_TO_BYTE := USINT_TO_BYTE(BYTE_TO_USINT(SHL(OCT_TO_BYTE,3)) + intX - 48);
    	END_IF
    	pt ACCESS (ADR(pt) + 1);
    END_FOR

    (* revision histroy
    hm	18. jun. 2008	rev 1.0
    	original release

    hm	20. sep. 2008	rev 1.1
    	changed length of input string from 20 to 10

    *)

END_FUNCTION

(* ---- OCT_TO_DWORD.st ---- *)
FUNCTION OCT_TO_DWORD
    (*http://www.oscat.de/images/OSCATBasic/oscat_basic333_en.pdf#page=176*)
    pt ACCESS ADR(OCT);
    stop := LEN(OCT);
    FOR i := 1 TO stop DO
    	(* read the first character and subtract 48 to get value in decimal 0 = 48 *)
    	X := pt;
        intX := BYTE_TO_USINT(X);
    	(* calculate the value of the digit *)
    	IF intX > 47 AND intX < 56 THEN
    		OCT_TO_DWORD := UDINT_TO_DWORD(DWORD_TO_UDINT(SHL(OCT_TO_DWORD,3)) + intX - 48);
    	END_IF
    	pt ACCESS (ADR(pt) + 1);
    END_FOR

    (* revision histroy
    hm	18. jun. 2008	rev 1.0
    	original release

    *)

END_FUNCTION

(* ---- OFFSET.st ---- *)
FUNCTION OFFSET
    (*http://www.oscat.de/images/OSCATBasic/oscat_basic333_en.pdf#page=282*)
    IF D THEN OFFSET := DEFAULT; ELSE OFFSET := X; END_IF
    IF O1 THEN OFFSET := OFFSET + OFFSET_1; END_IF
    IF O2 THEN OFFSET := OFFSET + OFFSET_2; END_IF
    IF O3 THEN OFFSET := OFFSET + OFFSET_3; END_IF
    IF O4 THEN OFFSET := OFFSET + OFFSET_4; END_IF

    (* revision history
    hm	12. jan 2007
    	original version

    *)
END_FUNCTION

(* ---- OFFSET2.st ---- *)
FUNCTION OFFSET2
    (*http://www.oscat.de/images/OSCATBasic/oscat_basic333_en.pdf#page=285*)
    IF D THEN OFFSET2 := DEFAULT; ELSE OFFSET2 := X; END_IF
    IF O4 THEN OFFSET2 := OFFSET2 + OFFSET_4;
    ELSIF O3 THEN OFFSET2 := OFFSET2 + OFFSET_3;
    ELSIF O2 THEN OFFSET2 := OFFSET2 + OFFSET_2;
    ELSIF O1 THEN OFFSET2 := OFFSET2 + OFFSET_1;
    END_IF
END_FUNCTION

(* ---- OM_TO_F.st ---- *)
FUNCTION OM_TO_F
    (*http://www.oscat.de/images/OSCATBasic/oscat_basic333_en.pdf#page=369*)
    OM_TO_F := OM / cPI2;

    (* revision history
    hm	22. jan. 2007	rev 1.0
    	original version

    hm	18. oct. 2008	rev 1.1
    	using math constants

    *)
END_FUNCTION

(* ---- OSCAT_VERSION.st ---- *)
FUNCTION OSCAT_VERSION
    (*http://www.oscat.de/images/OSCATBasic/oscat_basic333_en.pdf#page=37*)
    IF IN THEN
    	OSCAT_VERSION := DATE_TO_DWORD(D#2021-02-03);
    ELSE
    	OSCAT_VERSION := 334;
    END_IF

    (* revision history
    hm	6. oct 2006	rev 1.0
    	original version

    hm	16. dec 2007	rev 1.1
    	added possibility to return date and version depending on IN.

    *)
END_FUNCTION

(* ---- OVERRIDE.st ---- *)
FUNCTION OVERRIDE
    (*http://www.oscat.de/images/OSCATBasic/oscat_basic333_en.pdf#page=286*)
    IF E1 THEN OVERRIDE := X1; END_IF
    IF E2 AND ABS(X2) > ABS(OVERRIDE) THEN OVERRIDE := X2; END_IF
    IF E3 AND ABS(X3) > ABS(OVERRIDE) THEN OVERRIDE := X3; END_IF

    (* revision history
    hm	4.11.2007		rev 1.0
    	original version

    *)

END_FUNCTION

(* ---- PARITY.st ---- *)
FUNCTION PARITY
    (*http://www.oscat.de/images/OSCATBasic/oscat_basic333_en.pdf#page=230*)
    WHILE IN > 0 DO
    	PARITY := PARITY XOR IN.0 XOR IN.1 XOR IN.2 XOR IN.3;
    	IN := SHR(IN,4);
    END_WHILE

    (* code before rev 1.2
    WHILE IN > 0 DO
    	IF IN.0 THEN cnt := cnt +1; END_IF
    	IN := SHR(IN,1);
    END_WHILE
    IF (cnt MOD 2) = 1 THEN PARITY := TRUE; ELSE PARITY := FALSE; END_IF
    *)

    (* revision history

    rev 1.0 hm 1 sep 2006
    	original version

    rev 1.1 hm 10.9.2007
    	changed algorithm to improve performance

    rev 1.2	hm	8 dec 2007
    	changed algorithm to improve performance

    rev 1.3	hm	18 feb 2008
    	changed algorithm to improve performance
    *)
END_FUNCTION

(* ---- PERIOD.st ---- *)
FUNCTION PERIOD
    (*http://www.oscat.de/images/OSCATBasic/oscat_basic333_en.pdf#page=131*)
    day1 := DAY_OF_YEAR(D1);
    day2 := DAY_OF_YEAR(D2);
    dayx := DAY_OF_YEAR(DX);
    IF NOT LEAP_OF_DATE(DX) AND dayx > 58 THEN dayx := dayx + 1; END_IF
    IF NOT LEAP_OF_DATE(D1) AND day1 > 58 THEN day1 := day1 + 1; END_IF
    IF NOT LEAP_OF_DATE(D2) AND day2 > 58 THEN day2 := day2 + 1; END_IF

    IF day2 < day1 THEN
    	(* the PERIOD spans over the new year *)
    	PERIOD := dayx <= day2 OR dayx >= day1;
    ELSE
    	PERIOD := dayx >= day1 AND dayx <= day2;
    END_IF

    (* code before rev 1.2
    yx := year(DX);
    p1 := date_add(D1,0,0,0,yx - year(D1));
    p2 := date_add(D2,0,0,0,yx - year(D2));

    IF p2 >= p1 THEN
    	PERIOD := DX <= p2  AND DX >= p1;
    ELSE
    	PERIOD := DX <= p2 OR DX >= p1;
    END_IF
    *)

    (* revision history

    hm		19. sep 2007	rev 1.0
    	original version

    hm		20. sep 2007	rev 1.1
    	corrected a problem with leap year

    hm		4. jan 2008		rev 1.2
    	changed code for better performance

    hm		22. mar. 2008	rev 1.3
    	function would deliver wrong results when D1, D2 or DX are a leap_year

    *)
END_FUNCTION

(* ---- PERIOD2.st ---- *)
FUNCTION PERIOD2
    (*http://www.oscat.de/images/OSCATBasic/oscat_basic333_en.pdf#page=131*)
    PERIOD2 := 	(DX >= DP[0,0] AND DX <= DP[0,1]) OR
    			(DX >= DP[1,0] AND DX <= DP[1,1]) OR
    			(DX >= DP[2,0] AND DX <= DP[2,1]) OR
    			(DX >= DP[3,0] AND DX <= DP[3,1]);

    (* revision history

    hm		27. apr 2008	rev 1.0
    	original version

    *)
END_FUNCTION

(* ---- POLYNOM_INT.st ---- *)
FUNCTION POLYNOM_INT
    (*http://www.oscat.de/images/OSCATBasic/oscat_basic333_en.pdf#page=102*)
    (*make sure n is bound within the array size *)
    PTS := MIN(PTS, 5);

    (* this part is only to calculate the polynom parameters, which are then stores in the Y array
    	the array values, it is not needed during runtime, unless the parameters will change during runtime
    	the remaining code without this setup code can be used within a function to calculate specific functions
    	the content of the arrays is then used as constant values within the function *)

    FOR I := 1 TO PTS DO
    	stop := I + 1;
       	FOR J := PTS TO stop BY -1 DO
       		XY[J,1] := (XY[J,1] - XY[J-1,1]) / (XY[J,0] - XY[J-I,0]);
    	END_FOR
    END_FOR

    (* this part is the actual calculation *)
    POLYNOM_INT := 0.0;
    FOR I := PTS TO 1 BY -1 DO
           POLYNOM_INT := POLYNOM_INT * (X - XY[I,0]) + XY[I,1];
    END_FOR

    (* revision history
    hm	8. okt 2007	rev 1.0
    	original version

    hm	17. dec 2007	rev 1.1
    	init makes no sense for a function

    hm	22. feb 2008	rev 1.2
    	improved performance

    hm	10. mar. 2009	rev 1.3
    	changed syntax of real constants to 0.0

    *)
END_FUNCTION

(* ---- PT_TO_F.st ---- *)
FUNCTION PT_TO_F
    (*http://www.oscat.de/images/OSCATBasic/oscat_basic333_en.pdf#page=372*)
    PT_TO_F := 1000.0 / DWORD_TO_REAL(TIME_TO_DWORD(PT));

    (*	revision history
    hm	4. aug. 2006	rev 1.0
    	original version

    hm	11. mar. 2009	rev 1.1
    	real constants updated to new systax using dot

    *)

END_FUNCTION

(* ---- R2_ABS.st ---- *)
FUNCTION R2_ABS
    (*http://www.oscat.de/images/OSCATBasic/oscat_basic333_en.pdf#page=93*)
    IF X.RX >= 0.0 THEN
    	RETVAL.RX := X.RX;
    	RETVAL.R1 := X.R1;
    ELSE
    	RETVAL.RX := -X.RX;
    	RETVAL.R1 := -X.R1;
    END_IF
    R2_ABS:=TRUE;

    (* revision history
    hm	21. mar. 2008	rev 1.0
    	original version

    hm	10. mar. 2009 rev 1.1
    	real constants updated to new systax using dot

    *)
END_FUNCTION

(* ---- R2_ADD.st ---- *)
FUNCTION R2_ADD
    (*http://www.oscat.de/images/OSCATBasic/oscat_basic333_en.pdf#page=93*)
    temp := X.RX;
    RETVAL.RX := Y + X.R1 + X.RX;
    RETVAL.R1 := temp - RETVAL.RX + Y + X.R1;
    R2_ADD:=TRUE;

    (* revision history
    hm		20.3.2008	rev 1.0
    	original version

    *)
END_FUNCTION

(* ---- R2_ADD2.st ---- *)
FUNCTION R2_ADD2
    (*http://www.oscat.de/images/OSCATBasic/oscat_basic333_en.pdf#page=94*)
    RETVAL.R1 := X.R1 + Y.R1;
    RETVAL.RX := X.RX + Y.RX;
    R2_ADD2 := TRUE;

    (* revision history
    hm		20.3.2008	rev 1.0
    	original version

    *)
END_FUNCTION

(* ---- R2_MUL.st ---- *)
FUNCTION R2_MUL
    (*http://www.oscat.de/images/OSCATBasic/oscat_basic333_en.pdf#page=94*)
    RETVAL.RX := X.RX * Y;
    RETVAL.R1 := X.R1 * Y;
    R2_MUL:=TRUE;

    (* revision history
    hm		20.3.2008	rev 1.0
    	original version

    *)
END_FUNCTION

(* ---- R2_SET.st ---- *)
FUNCTION R2_SET
    (*http://www.oscat.de/images/OSCATBasic/oscat_basic333_en.pdf#page=95*)
    RETVAL.RX := X;
    RETVAL.R1 := 0.0;
    R2_SET:=TRUE;

    (* revision history
    hm	2. jun. 2008	rev 1.0
    	original version

    hm	10. mar. 2009	rev 1.1
    	real constants updated to new systax using dot

    *)
END_FUNCTION

(* ---- RAD.st ---- *)
FUNCTION RAD
    (*http://www.oscat.de/images/OSCATBasic/oscat_basic333_en.pdf#page=61*)
    RAD := MODR(0.0174532925199433 * DEG, cPI2);

    (* revision history
    hm	4. aug 2006		rev 1.0
    	original version

    hm 	16. oct 2007	rev 1.1
    	added modr statement which prohibits RAD to become bigger than 2PI

    hm	18. oct 2008	rev 1.2
    	using math constants

    *)
END_FUNCTION

(* ---- RANGE_TO_BYTE.st ---- *)
FUNCTION RANGE_TO_BYTE
    (*http://www.oscat.de/images/OSCATBasic/oscat_basic333_en.pdf#page=288*)
    RANGE_TO_BYTE := INT_TO_BYTE(DINT_TO_INT(TRUNC((LIMIT(LOW, X, HIGH) - LOW) * 255.0 / (HIGH - LOW))));

    (* revision history
    hm	9. jan 2008		rev 1.0
    	original version

    *)

END_FUNCTION

(* ---- RANGE_TO_WORD.st ---- *)
FUNCTION RANGE_TO_WORD
    (*http://www.oscat.de/images/OSCATBasic/oscat_basic333_en.pdf#page=288*)
    RANGE_TO_WORD := DINT_TO_WORD(TRUNC((LIMIT(LOW,X,HIGH)-LOW) * 65535.0 / (HIGH - LOW)));

    (* revision history
    hm	9. jan 2008		rev 1.0
    	original version

    *)

END_FUNCTION

(* ---- RDM.st ---- *)
FUNCTION RDM
    (*http://www.oscat.de/images/OSCATBasic/oscat_basic333_en.pdf#page=62*)
    tn := T_PLC_MS();
    tc := BIT_COUNT(UDINT_TO_DWORD(tn));
    tn.31 := tn.2;
    tn.30 := tn.5;
    tn.29 := tn.4;
    tn.28 := tn.1;
    tn.27 := tn.0;
    tn.26 := tn.7;
    tn.25 := tn.6;
    tn.24 := tn.3;
    tn := ROL(tn,BIT_COUNT(UDINT_TO_DWORD(tn))) OR 16#80000001;
    tn := tn MOD 71474513 + INT_TO_UDINT(tc + 77);
    RDM := FRACT(UDINT_TO_REAL(tn) / 10000000.0 * (ce - LIMIT(0.0,LAST,1.0)));

    (*
    pt := ADR(temp);
    pt := (T_PLC_MS() AND 16#007FFFFF) OR 16#3D000000;
    RDM := fract(modR(temp*e+pi1, PI1-LAST) + modR(temp*PI1+e + LAST,e-LAST));
    *)

    (* revision history
    hm		16. jan 2007		rev 1.0
    	original version

    hm		11. nov 2007		rev 1.1
    	changed time() into t_plc_ms()

    hm		20. nov 2007		rev 1.2
    	changed code of temp calculation to avoid overflow in modr due to resuclt would not fit DINT for high timeer values

    hm		5. jan 2008		rev 1.3
    	changed calculation of temp to avoid problem with high values of t_plc_ms

    hm		2. feb 2008		rev 1.4
    	changed algorithm to avoind non iec functions and guarantee more randomness

    hm	10. mar. 2008		rev 1.5
    	make sure LAST will be between 0 and 1 to avoid invalid results

    hm	16. mar. 2008		rev 1.6
    	added conversion for tc to avoid warnings under codesys 3.0

    hm	18. may. 2008		rev 1.7
    	changed constant E to E1

    hm	18. oct. 2008		rev 1.8
    	using math constants

    hm	10. mar. 2009		rev 1.9
    	real constants updated to new systax using dot

    *)
END_FUNCTION

(* ---- RDM2.st ---- *)
FUNCTION RDM2
    (*http://www.oscat.de/images/OSCATBasic/oscat_basic333_en.pdf#page=62*)
    RDM2 := DINT_TO_INT(TRUNC(RDM(FRACT(LAST * cPI)) * (HIGH - LOW + 1)) + LOW);

    (* revision history
    hm		29. feb 2008		rev 1.0
    	original version

    hm		18. oct. 2008		rev 1.1
    	using math constants

    *)
END_FUNCTION

(* ---- RDMDW.st ---- *)
FUNCTION RDMDW
    (*http://www.oscat.de/images/OSCATBasic/oscat_basic333_en.pdf#page=63*)
    M := BIT_COUNT(LAST);
    RX := RDM(FRACT(M * cPI));
    RDMDW := SHL(REAL_TO_DWORD(RX*65535),16);
    RX := RDM(FRACT(M * ce));
    RDMDW := RDMDW OR (REAL_TO_DWORD(RX*65535) AND 16#0000FFFF);

    (* revision history
    hm		14. mar 2008		rev 1.0
    	original version

    hm		18. may. 2008		rev 1.1
    	changed constant E to E1

    hm		18. oct. 2008		rev 1.2
    	using math constants

    *)
END_FUNCTION

(* ---- REAL_TO_DW.st ---- *)
FUNCTION REAL_TO_DW
    (*http://www.oscat.de/images/OSCATBasic/oscat_basic333_en.pdf#page=231*)
    pt ACCESS ADR(X);
    REAL_TO_DW := pt;

    (* revision history
    hm	18. apr. 2008
    	original version

    *)
END_FUNCTION

(* ---- REAL_TO_FRAC.st ---- *)
FUNCTION REAL_TO_FRAC
    (*http://www.oscat.de/images/OSCATBasic/oscat_basic333_en.pdf#page=64*)
    IF X < 0.0 THEN
    	sign := TRUE;								(* Vorzeichen merken *)
    	X := ABS(X);								(* Absolutwert berechnen *)
    END_IF

    REPEAT
    	X_gerundet := REAL_TO_DINT(X);

    	(* Zaehler berechnen *)
    	temp := Numerator * X_gerundet + Numerator_old;		(* Zaehler um Vorkammawert erweitern *)
    	Numerator_old := Numerator;							(* Zaehler der letzten Berechnung speichern *)
    	Numerator := temp;									(* Zaehler dieser Berechnung speichern *)

    	(* Nenner berechnen *)
    	temp := Denominator * X_gerundet + Denominator_old;	(* Nenner um Vorkammawert erweitern *)
    	Denominator_old := Denominator;						(* Nenner der letzten Berechnung speichern *)
    	Denominator := temp;								(* Nenner dieser Berechnung speichern *)

    	(* Restwert berechnen *)
    	X_ohne_Nachkomma := DINT_TO_REAL(X_gerundet);
    	IF X = X_ohne_Nachkomma THEN						(* Bruch geht ohne Rest auf *)
    		IF ABS(Denominator) <= N THEN						(* kein Rundungsfehler *)
    			Numerator_old := Numerator;					(* Numerator_old wird von Funktion zurückgegeben *)
    			Denominator_old := Denominator;			(* Denominator_old wird von Funktion zurückgegeben *)
    		END_IF
    		EXIT;											(* keine weitere Berechnung notwendig *)
    	ELSE
    		X := 1.0 / (X - X_ohne_Nachkomma);				(* Kehrwert vom Rest -> Neuer Bruch *)
    	END_IF

    UNTIL
    	ABS(Denominator) > N
    END_REPEAT

    (* correct sign if X was negative *)
    IF sign THEN
    	RETVAL.NUMERATOR := -1 * ABS(DINT_TO_INT(Numerator_old));
    ELSE
    	RETVAL.NUMERATOR :=  ABS(DINT_TO_INT(Numerator_old));
    END_IF
    RETVAL.DENOMINATOR := ABS(DINT_TO_INT(Denominator_old));
    REAL_TO_FRAC:=TRUE;

    (* revision history
    hm		19. jan. 2011	rev 1.0
    	original version

    ad		06. apr. 2011	rev 1.1
    	optimized code
    *)
END_FUNCTION

(* ---- REAL_TO_STRF.st ---- *)
FUNCTION REAL_TO_STRF
    (*http://www.oscat.de/images/OSCATBasic/oscat_basic333_en.pdf#page=176*)
    (* LIMIT N to 0 .. 7 *)
    N := LIMIT(0,N,7);
    (* round the input to N digits and convert to string *)
    O := ABS(IN) * EXP10(N);
    RETVAL := DINT_TO_STRING(REAL_TO_DINT(O));
    (* add zeroes IN front to make sure sting is at least 8 digits long *)
    FOR i := LEN(RETVAL) TO N DO RETVAL := CONCAT('0', RETVAL); END_FOR
    (* add a dot if N > 0 *)
    IF N > 0 THEN RETVAL := INSERT(RETVAL, D, LEN(RETVAL) - N); END_IF
    (* add a minus sign if IN is negative *)
    IF IN < 0 THEN RETVAL := CONCAT('-', RETVAL); END_IF
    REAL_TO_STRF := TRUE;

    (* revision history
    hm	26 jan 2007	rev 1.0
    	original version

    hm	20. nov. 2007	rev 1.1
    	when N=0 ther will be no dot at the end of the string.

    hm	15. dec. 2007	rev 1.2
    	changed code for better performance

    hm	4. mar. 2008	rev 1.3
    	result is now rounded instead of trunc

    hm	20. mar. 2008	rev 1.4
    	changed trunc to real_to_dint because trunc was generating wrong values on wago 842

    hm	29. mar. 2008	rev 1.5
    	changed STRING to STRING(20)

    hm	4. apr. 2008	rev 1.6
    	added variable O to avoid an error uner CoDeSys SP PLCWinNT V2.4

    hm	27. feb. 2009	rev 1.7
    	added a missing zero for IN < 1

    hm 2. jan 2012	rev 1.8
    	added input parameter D to specify decimal separator
    *)

END_FUNCTION

(* ---- REFLECT.st ---- *)
FUNCTION REFLECT
    (*http://www.oscat.de/images/OSCATBasic/oscat_basic333_en.pdf#page=232*)
    REFLECT := 0;
    FOR i := 1 TO L DO
    	REFLECT := SHL(REFLECT, 1) OR BOOL_TO_DWORD(D.0);
    	D := SHR(D, 1);
    END_FOR
    REFLECT := REFLECT OR SHL(D, L);

    (* revision history
    hm	 16. jan 2011
    	new module

    *)
END_FUNCTION

(* ---- REFRACTION.st ---- *)
FUNCTION REFRACTION
    (*http://www.oscat.de/images/OSCATBasic/oscat_basic333_en.pdf#page=132*)
    ELEV := LIMIT(-1.9, ELEV, 80.0);
    REFRACTION := 0.0174532925199433 / TAN(0.0174532925199433 * (ELEV + 10.3 / (ELEV + 5.11)));

    (* revision histroy
    hm	14. jul. 2008	rev 1.0
    	original release

    hm	7. mar. 2009	rev 1.1
    	using new formula

    *)

END_FUNCTION

(* ---- REPLACE_ALL.st ---- *)
FUNCTION REPLACE_ALL
    (*http://www.oscat.de/images/OSCATBasic/oscat_basic333_en.pdf#page=177*)
    RETVAL := STR;
    lx := LEN(SRC);
    lp := LEN(REP);
    pos := FINDP(RETVAL, SRC, 1);
    WHILE pos > 0 DO
    	RETVAL := REPLACE(RETVAL,REP,lx, pos);
    	pos := FINDP(RETVAL, SRC, pos + lp);
    END_WHILE
    REPLACE_ALL := TRUE;
    (* revision histroy
    hm	4. feb. 2008	rev 1.0
    	original release

    hm	29. mar. 2008	rev 1.1
    	changed STRING to STRING(STRING_LENGTH)
    *)

END_FUNCTION

(* ---- REPLACE_CHARS.st ---- *)
FUNCTION REPLACE_CHARS
    (*http://www.oscat.de/images/OSCATBasic/oscat_basic333_en.pdf#page=177*)
    RETVAL := STR;
    (* make sure REP and SRC are of same length and length is > 0 *)
    a := LEN(SRC);
    b := LEN(REP);
    IF a < b THEN
    	REP := LEFT(REP, a);
    ELSIF b < a THEN
    	SRC := LEFT(SRC, b);
    END_IF

    (* search the string and replace if necessary *)
    stp := LEN(STR);
    FOR a := 1 TO stp DO
    	c := MID(RETVAL, 1, a);
    	b := FIND(SRC, c);
    	IF b > 0 THEN
    		RETVAL := REPLACE(RETVAL, MID(REP, 1, b), 1, a);
    	END_IF
    END_FOR
    REPLACE_CHARS := TRUE;

    (* revision history
    hm	14. may. 2008	rev 1.0
    	original version

    *)

END_FUNCTION

(* ---- REPLACE_UML.st ---- *)
FUNCTION REPLACE_UML
    (*http://www.oscat.de/images/OSCATBasic/oscat_basic333_en.pdf#page=178*)
    pt ACCESS ADR(STR);
    pto ACCESS ADR(RETVAL);
    ptm ACCESS (ADR(pto) + INT_TO_UDINT(STRING_LENGTH));
    pt1 ACCESS ADR(su);
    pt2 ACCESS (ADR(pt1) + 1);
    L := LEN(STR);
    WHILE pos < L AND pos < STRING_LENGTH DO
    	IF pt < 127 THEN
    		(* no uml character simlply copy the character*)
    		pto := pt;
    	ELSE
    		(* convert the uml character *)
    		TO_UML(pt, su);
    		(* we must make sure pointer are not out of range *)
    		pto := pt1;
    		IF ADR(pto) < ADR(ptm) AND pt2 > 0 THEN
    			pto ACCESS (ADR(pto) + 1);
    			pto := pt2;
    		END_IF
    	END_IF
    	(* increment pointers *)
    	pt ACCESS (ADR(pt) + 1);
    	pto ACCESS (ADR(pto) + 1);
    	pos := pos + 1;
    END_WHILE

    (* properly close the output string *)
    pto := 0;
    REPLACE_UML := TRUE;

    (* revision history
    hm	29. feb 2008	rev 1.0
    	original version

    hm	29. mar. 2008	rev 1.1
    	changed STRING to STRING(STRING_LENGHT)
    	new code to avoid pointer out of range
    	use new function to_uml
    *)
END_FUNCTION

(* ---- RES_NI.st ---- *)
FUNCTION RES_NI
    (*http://www.oscat.de/images/OSCATBasic/oscat_basic333_en.pdf#page=318*)
    T2 := T * T;
    RES_NI := R0 + A * T + B * T2 + C * T2 * T2;

    (* revision history

    hm	4.8.2006		rev 1.0
    	original version

    hm	13.9.2007		rev 1.1
    	changed coding for better performance

    hm	2. dec. 2007	rev 1.2
    	changed code for better performance
    *)

    (*

     Auszug aus DIN 43760 für Ni100

    °C		R		°C		R		°C	R		°C		R		°C		R

    -60 	69,5 	-10 	94,6 	40 	123,0 	90 		154,9 	140 	190,9
    -55 	71,9 	-5 		97,3 	45 	126,0 	95 		158,3 	145 	194,8
    -50 	74,3 	0 		100,0 	50 	129,1 	100 	161,8 	150 	198,7
    -45 	76,7 	5 		102,8 	55 	132,2 	105 	165,3 	155 	202,6
    -40 	79,1 	10 		105,6 	60 	135,3 	110 	168,8 	160 	206,6
    -35 	81,6 	15 		108,4 	65 	138,5 	115 	172,4 	165 	210,7
    -30 	84,2 	20 		111,2 	70 	141,7 	120 	176,0 	170 	214,8
    -25 	86,7 	25 		114,1 	75 	145,0 	125 	179,6 	175 	219,0
    -20 	89,3 	30 		117,1 	80 	148,3 	130 	183,3 	180 	223,2
    -15 	91,9 	35 		120,0 	85 	151,6 	135 	187,1

    *)
END_FUNCTION

(* ---- RES_NTC.st ---- *)
FUNCTION RES_NTC
    (*http://www.oscat.de/images/OSCATBasic/oscat_basic333_en.pdf#page=319*)
    RES_NTC := RN * EXP(B * (1.0 / (T+273.15) - 0.00335401643468053));

    (* revision history

    hm 30. dec. 2008	rev 1.0
    	original version

    hm	11. mar. 2009	rev 1.1
    	changed real constants to use dot syntax

    *)
END_FUNCTION

(* ---- RES_PT.st ---- *)
FUNCTION RES_PT
    (*http://www.oscat.de/images/OSCATBasic/oscat_basic333_en.pdf#page=322*)
    T2 := T * T;

    IF T >= 0.0 THEN
    	RES_PT := R0 * ( 1.0 + A * T + B * T2);
    ELSE
    	RES_PT := R0 * ( 1.0 + A * T + B * T2 + C * (T - 100.0) * T2 * T);
    END_IF

    (* revision history
    hm	4. aug. 2006	rev 1.1
    	original version

    hm	2. dec 2007	rev 1.2
    	changed code for better performance

    hm	11. mar. 2009	rev 1.3
    	changed real constants to use dot syntax

    *)

    (*
     Auszug aus DIN 43760 für Pt100

    °C		R		°C		R		°C	R			°C		R			°C		R			°C		R

    -200 	18,49 	-100 	60,25 	0 	100,00 	100 	138,50 	200 	175,84 	300 	212,02
    -195 	20,65 	-95 	62,28 	5 	101,95 	105 	140,39 	205 	177,68 	305 	213,80
    -190 	22,80 	-90 	64,30 	10 	103,90 	110 	142,29 	210 	179,51 	310 	215,57
    -185 	24,94 	-85 	66,31 	15 	105,85 	115 	144,17 	215 	181,34 	315 	217,35
    -180 	27,08 	-80 	68,33 	20 	107,79 	120 	146,06 	220 	183,17 	320 	219,12
    -175 	29,20 	-75 	70,33 	25 	109,73 	125 	147,94 	225 	184,99 	325 	220,88
    -170 	31,32 	-70 	72,33 	30 	111,67 	130 	149,82 	230 	186,82 	330 	222,65
    -165 	33,43 	-65 	74,33 	35 	113,61 	135 	151,70 	235 	188,63 	335 	224,41
    -160 	35,33 	-60 	76,33 	40 	115,54 	140 	153,58 	240 	190,45 	340 	226,17
    -155 	37,63 	-55 	78,32 	45 	117,47 	145 	155,45 	245 	192,26 	345 	227,92
    -150 	39,71 	-50 	80,31 	50 	119,40 	150 	157,31 	250 	194,07 	350 	229,67
    -145 	41,79 	-45 	82,29 	55 	121,32 	155 	159,18 	255 	195,88 	355 	231,42
    -140 	43,87 	-40 	84,27 	60 	123,24 	160 	161,04 	260 	197,69 	360 	233,17
    -135 	45,94 	-35 	86,25 	65 	125,16 	165 	162,90 	265 	199,49 	365 	234,91
    -130 	48,00 	-30 	88,22 	70 	127,07 	170 	164,76 	270 	201,29 	370 	236,65
    -125 	50,06 	-25 	90,19 	75 	128,98 	175 	166,61 	275 	203,08 	375 	238,39
    -120 	52,11 	-20 	92,16 	80 	130,89 	180 	168,46 	280 	204,88 	380 	240,13
    -115 	54,15 	-15 	94,12 	85 	132,80 	185 	170,31 	285 	206,67 	385 	241,86
    -110 	56,19 	-10 	96,09 	90 	134,70 	190 	172,16 	290 	208,45 	390 	243,59
    -105 	58,22 	-5 		98,04 	95 	136,60 	195 	174,00 	295 	210,24 	395 	245,31

    *)
    (*
    revision history

    *)
END_FUNCTION

(* ---- RES_SI.st ---- *)
FUNCTION RES_SI
    (*http://www.oscat.de/images/OSCATBasic/oscat_basic333_en.pdf#page=323*)
    TX := T - TS;
    RES_SI := RS * ( 1.0 + A * TX + B * TX * TX);

    (* revision history
    hm	4. aug 2006	rev 1.0
    	original version

    hm	2. dec 2007	rev 1.1
    	changed code for better performance

    hm	11. mar. 2009	rev 1.2
    	changed real constants to use dot syntax

    *)
END_FUNCTION
